// TIA Portal project "Can_Van_An_Modbus_ASCII" (V21)

(* hardware
DEVICE "S7-1500/ET200MP station_1"  S7-1500 station
   slot 0: "Rail_0"  Rack  6ES7 590-1***0-0AA0
   slot 1: "PLC_1"  CPU 1513-1 PN  6ES7 513-1AL02-0AB0  V2.9
      slot 3: "CPU display_1"  6ES7591-1AA00-0AA0
      slot 32768: "PROFINET interface_1"  X1
         slot 32769: "Port_1"  X1 P1
         slot 32770: "Port_2"  X1 P2
      slot 34817: "Virtual CP interface port_1"  Virtual CP interface port  Virtual CP interface port
DEVICE "ET 200SP station_1"  ET 200SP-Station
   slot 0: "Rack_0"  Rack  6ES5 710-8MAx1
   slot 0: "IO device_1"  IM 155-6 PN ST  6ES7 155-6AU01-0BN0  V4.2
   slot 1: "CM PtP_1"  CM PtP  6ES7 137-6AA01-0BA0  V2.0
      slot 1: "CM PtP_1"  CM PtP Sub
   slot 2: "Server module_1"  Server module  6ES7 193-6PA00-0AA0  V1.1
      slot 1: "Server module_1"  Server module
   slot 127: "BA 2xRJ45"  BA 2xRJ45  6ES7 193-6AR00-0AA0  V0.0
      slot 1: "Port_1"  X1 P1R  6ES7 193-6AR00-0AA0  V0.0
      slot 2: "Port_2"  X1 P2R  6ES7 193-6AR00-0AA0  V0.0
*)

// ===== PLC "PLC_1"  CPU 1513-1 PN =====

VAR_GLOBAL   // PLC tag table "1_Default tag table"
   "System_Byte" AT %MB1 : Byte;
   "FirstScan" AT %M1.0 : Bool;
   "DiagStatusUpdate" AT %M1.1 : Bool;
   "AlwaysTRUE" AT %M1.2 : Bool;
   "AlwaysFALSE" AT %M1.3 : Bool;
   "Clock_Byte" AT %MB0 : Byte;
   "Clock_10Hz" AT %M0.0 : Bool;
   "Clock_5Hz" AT %M0.1 : Bool;
   "Clock_2.5Hz" AT %M0.2 : Bool;
   "Clock_2Hz" AT %M0.3 : Bool;
   "Clock_1.25Hz" AT %M0.4 : Bool;
   "Clock_1Hz" AT %M0.5 : Bool;
   "Clock_0.625Hz" AT %M0.6 : Bool;
   "Clock_0.5Hz" AT %M0.7 : Bool;
END_VAR

VAR_GLOBAL   // PLC tag table "2_Bit_Tam(2-10)"
   "bTrigger1" AT %M2.0 : Bool;
   "bTrigger2" AT %M2.1 : Bool;
   "bTrigger3" AT %M2.2 : Bool;
   "bTrigger4" AT %M2.3 : Bool;
   "bTrigger5" AT %M2.4 : Bool;
   "bTrigger6" AT %M2.5 : Bool;
   "bTrigger7" AT %M2.6 : Bool;
   "bTrigger8" AT %M2.7 : Bool;
   "bTrigger9" AT %M3.0 : Bool;
   "bTrigger10" AT %M3.1 : Bool;
END_VAR

VAR_GLOBAL   // PLC tag table "3_DataNodeRed(100-200)"
   "diWeight" AT %MD100 : DInt;
   "wErrorCodeWeight" AT %MW104 : Word;
   "wStatusPLC" AT %MW106 : Word;
END_VAR

TYPE "typePortConfigSettings"
   STRUCT
      port : Int;
      protocol : Int;
      baud : Int;
      parity : Int;
      dataBis : Int;
      stopBits : Int;
      flowCntr : Int;
   END_STRUCT;
END_TYPE

TYPE "StartConditionReceive"
   STRUCT
      wStartCond : Word;
      wIdleTime : Word;
      StartChar : Byte;
   END_STRUCT;
END_TYPE

// folder: Common

TYPE "typeDiagnostics"
TITLE = typeDiagnostics
// Provides a structure for detailed diagnostics
   STRUCT
      status : Word;   // Status of the block or error identification when error occurred
      subfunctionStatus : DWord;   // Status or return value of called FBs, FCs and system blocks
      stateNumber : DInt;   // State in the state machine of the block where the error occurred
   END_STRUCT;
END_TYPE

// folder: LMQTT

TYPE "LMQTT_typeConnParam"
TITLE = LMQTT_typeConnParams
// Specifies connection parameters for the mqtt connection
   STRUCT
      hwId : Hw_Any;   // Hardware identifier of the interface. 0: interface is selected automatically
      connId : Conn_Ouc := 1;   // Unique connection identifier (1..4095)
      broker : String;   // Hostname or IP address of broker
      port : UInt := 1883;   // Port on the broker
      tls : Struct   // Parameters for TLS encryption
         enableTls : Bool;   // TRUE: Enables TLS, FALSE: disable TLS
         validateServerIdentity : Bool;   // TRUE: Validate server certificate, FALSE: No validation of server certificate
         brokerCert : UDInt;   // ID of the broker's certificate in TIA Portal
         clientCert : UDInt;   // ID of the client's certificate in TIA Portal
      END_STRUCT;
      keepAlive : UInt;   // Keepalive mechanism for MQTT in seconds. 0: disabled.
   END_STRUCT;
END_TYPE

// folder: typeDefinitions

TYPE "LModbusAscii_typeAsciiConfiguration"
TITLE = Parameter dataset to configure Modbus interface
// Parameter dataset to configure Modbus interface
   STRUCT
      baud : UInt := 6;   // Baud rate, default is 9600 (6), 19200 (7), see manual for other definitions
      parity : UInt := 2;   // Parity, default is even (2), odd (3) or none (1)
      modeInterfacePTP : USInt := 4;   // Serial interface mode, default is RS485 (4, Half duplex, two-wire mode), RS232 (0, FullDuplex)
      numberOfRetries : USInt := 3;   // Number of retries if a transmission error occurs, default is 3
      transmissionWatchdog : Time := T#5S;   // Response timeout duration, default is 5 s
   END_STRUCT;
END_TYPE

TYPE "LModbusAscii_typeDiagnostics"
TITLE = typeDiagnosticsTemplate
   STRUCT
      status : Word;   // Status of the block or error identification when error occurred
      stateNumber : DInt;   // State in the state machine of the block where the error occurred
      subFunctionStatus : Word;   // Status or return value of called FBs, FCs and system blocks
   END_STRUCT;
END_TYPE

// folder: (top level)

DATA_BLOCK "Data_StateSystem"   // DB1
{ S7_Optimized_Access := 'FALSE' }
VERSION : 0.1
   VAR
      "LED_PLC-S7-1500" : Struct
         "PLC-S7-1500" : Hw_Io := 50;
         Mode : Int := 1;
         Ret_Val : Word;
      END_STRUCT;
      ET200SP : Struct
         Device1 : Array[0..127] of Bool;
         RetVal : Int;
      END_STRUCT;
      bPLC_OFF : Bool;
      bPLC_Run : Bool;
      bPLC_Stop : Bool;
      bESP200_OK : Bool;
      bESP200_Fault : Bool;
      bESP200_LostConnect : Bool;
      bDonePortConfig : Bool;
      bErrorPortConfig : Bool;
      wStatusPortConfig : Word;
      "bDoneSend Config" : Bool;
      bErrorSendConfig : Bool;
      wStatusSendConfig : Word;
      bDoneReceiveConfig : Bool;
      bErrorReceiveConfig : Bool;
      wStatusReceiveConfig : Word;
      bDoneModbusKeli : Bool;
      bBusyModbusKeli : Bool;
      bErrorModbuskeli : Bool;
      ConditionReceive : Receive_Conditions;
   END_VAR
BEGIN
END_DATA_BLOCK

DATA_BLOCK "LMQTT_Client_EMQX_DB"   // DB2
{ S7_Optimized_Access := 'TRUE' }
AUTHOR : Siemens Industry Online Support
FAMILY : LMQTT
VERSION : 4.2
// stored: InstanceOfName LMQTT_Client
"LMQTT_Client"
BEGIN
END_DATA_BLOCK

DATA_BLOCK "KELI_ReadWeight_DB"   // DB3
{ S7_Optimized_Access := 'TRUE' }
VERSION : 1.0
// stored: InstanceOfName KELI_ReadWeight
"KELI_ReadWeight"
BEGIN
END_DATA_BLOCK

DATA_BLOCK "MQTT_Client"   // DB5
{ S7_Optimized_Access := 'FALSE' }
VERSION : 0.1
   VAR
      Inputs : Struct
         enable : Bool;
         publish : Bool;
         subscribe : Bool;
         unsubscribe : Bool;
         connParam : "LMQTT_typeConnParam";
         cleanSession : Bool;
         clientIdentifier : WString;
         username : WString;
         password : WString;
         willtopic : WString;
         willMsgLen : UInt;
         qos : USInt;
         retain : Bool;
         mqttTopic : WString;
         publishMsgLen : UDInt;
         timeOut : Time;
      END_STRUCT;
      Outputs : Struct
         valid : Bool;
         done : Bool;
         busy : Bool;
         error : Bool;
         status : Word;
         diagnostics : "typeDiagnostics";
         sessionPresent : Bool;
         receivedMsgStatus : USInt;
         receivedMsgDataLen : UDInt;
      END_STRUCT;
      InOut : Struct
         willMsgPayload : Array[0..7] of Byte;
         publishMsgPayload : Array[0..7] of Byte;
         receivedTopic : WString;
         receivedMsgPayload : Array[0..7] of Byte;
      END_STRUCT;
   END_VAR
BEGIN
   Inputs.connParam.hwId := 64;
END_DATA_BLOCK

DATA_BLOCK "Data_Server"   // DB11
{ S7_Optimized_Access := 'FALSE' }
VERSION : 0.1
   VAR
      MB_TCPIP : TCON_IP_v4;
   END_VAR
BEGIN
   MB_TCPIP.InterfaceId := 64;
   MB_TCPIP.ID := 1;
   MB_TCPIP.ConnectionType := 11;
   MB_TCPIP.ActiveEstablished := False;
   MB_TCPIP.RemoteAddress.ADDR[1] := 0;
   MB_TCPIP.RemoteAddress.ADDR[2] := 0;
   MB_TCPIP.RemoteAddress.ADDR[3] := 0;
   MB_TCPIP.RemoteAddress.ADDR[4] := 0;
   MB_TCPIP.RemotePort := 0;
   MB_TCPIP.LocalPort := 502;
END_DATA_BLOCK

DATA_BLOCK "Data_FrameKeli"   // DB13
{ S7_Optimized_Access := 'FALSE' }
VERSION : 0.1
   VAR
      ton : TON_TIME;
      WeightRAW_RX : String;
      ReadWeight_TX : Array[0..7] of Byte;
   END_VAR
BEGIN
   ReadWeight_TX[1] := 16#03;   // function
   ReadWeight_TX[0] := 16#02;   // address
   ReadWeight_TX[3] := 16#01;   // Thanh ghi băt đầu low
   ReadWeight_TX[2] := 16#00;   // Thanh ghi băt đầu high
   ReadWeight_TX[4] := 16#00;   // Thanh ghi kết thúc high
   ReadWeight_TX[5] := 16#04;   // Thanh ghi kết thúc low
   ReadWeight_TX[6] := 16#15;   // CRC16L
   ReadWeight_TX[7] := 16#FA;   // CRC16L
END_DATA_BLOCK

FUNCTION_BLOCK "KELI_ReadWeight"   // FB3, SCL
{ S7_Optimized_Access := 'TRUE' }
VERSION : 1.1
// ===============================================================================
//  KELI_ReadWeight - Đọc khối lượng GROSS của đầu cân KELI D2008 qua MODBUS (TF = 1)
//  PLC: S7-1200 / S7-1500 + module CM RS485 (Freeport, dùng Send_P2P / Receive_P2P)
// -------------------------------------------------------------------------------
//  CÀI ĐẶT ĐẦU CÂN: tF = 1 (MODBUS command), Adr = địa chỉ 1..247, bt = baudrate, jn = parity
//  CÀI ĐẶT CỔNG CM (Port configuration):
//    - Baudrate / parity / 8 data bit / 1 stop bit: giống đầu cân
//    - Message end (Receive): "Recognize end of message by line idle time"
//      (đầu cân nghỉ >= 4 ký tự sau mỗi khung -> CM báo đã nhận đủ khung)
// 
//  KHUNG TIN (theo manual D2008, mục MODBUS command mode):
//    Lệnh gửi (requestFrame, 8 byte):
//      [0] địa chỉ  [1] 16#03  [2] 16#00  [3] 16#01  [4] 16#00  [5] 16#04  [6] CRC low  [7] CRC high
//      ví dụ địa chỉ 1: 16#01 03 00 01 00 04 15 C9
//    Phản hồi bình thường (13 byte):
//      [0] địa chỉ  [1] 16#03  [2] 16#08 (= 8 byte dữ liệu)
//      [3] dấu: '0' (16#30) = dương, '-' = âm  [4..9] 6 chữ số ASCII (Data5..Data0)  [10] số chữ số thập phân
//      [11] CRC low  [12] CRC high
//      ví dụ 20.00 kg: '0' '0' '0' '2' '0' '0' '0' '2' -> weight = 2000, decimals = 2
//    Phản hồi lỗi (exception, 5 byte): [0] địa chỉ  [1] 16#83  [2] mã exception  [3] CRC L  [4] CRC H
// 
//  CRC16 MODBUS: giá trị đầu 16#FFFF, đa thức 16#A001, tính trên mọi byte trừ 2 byte CRC,
//    gửi byte thấp trước, byte cao sau.
// 
//  OUTPUT GIÁ TRỊ CÂN:
//    weight    : khối lượng dạng số nguyên, có dấu, KHÔNG có dấu thập phân (vd 2000)
//    decimals  : số chữ số sau dấu thập phân (vd 2  ->  khối lượng thật = 2000 / 10^2 = 20.00)
//    weightRaw : chuỗi 8 ký tự đầu cân gửi về, đúng nguyên bản (vd '00020002')
// 
//  status : 0 = BAD (lỗi), 1 = GOOD (đọc tốt), 2 = UNCERTAIN (chưa có giá trị / đang retry)
// 
//  TỰ KHỞI ĐỘNG LẠI: autoRestart = TRUE -> sau khi báo lỗi, FB chờ restartDelay rồi
//    tự chạy lại từ đầu, không cần sườn lên ở execute. restartCount đếm số lần tự chạy lại.
//    resetRestartCount (IN_OUT): SCADA/HMI ghi TRUE -> restartCount = 0, FB tự trả tag về FALSE.
//      Nối vào 1 tag Bool trong DB (vd "HMI".resetRestartCount_Can1), không nối hằng số.
// 
//  [V1.1] ĐO THỜI GIAN PHẢN HỒI CỦA ĐẦU CÂN (timer độ phân giải 1 ms):
//    Bắt đầu đếm : khi FB bắt đầu gửi lệnh xuống đầu cân (vào bước 20 - SEND)
//    Kết thúc    : khi CM báo đã nhận xong khung trả lời (Receive_P2P.NDR ở bước 30)
//    KHÔNG tính  : thời gian kiểm tra CRC và đổi ra số cân (bước 40)
//    responseTime   : kết quả dạng Time (vd T#45MS)
//    responseTimeMs : kết quả dạng số ms (vd 45) - tiện hiển thị trên HMI / SCADA
//    Chỉ cập nhật khi nhận được khung; timeout / lỗi gửi -> giữ giá trị lần đo gần nhất.
//    Mỗi lần retry đo lại từ đầu -> kết quả là thời gian của lần gửi nhận được trả lời.
//    Lưu ý: FB chỉ thấy NDR khi được gọi, nên kết quả có thể lớn hơn thực tế tối đa 1 chu kỳ quét.
// 
//  BẢNG MÃ LỖI (errorCode) - subStatus cho biết thêm chi tiết:
//    16#0000 ERR_NONE                không lỗi
//    16#8101 ERR_PARAM_ADDRESS       requestFrame[0] không thuộc 1..247   sub = địa chỉ nhập
//    16#8102 ERR_PARAM_FUNCTION      requestFrame[1] khác 16#03            sub = mã nhập
//    16#8103 ERR_PARAM_REGISTER      thanh ghi khác 16#0001 (gross)        sub = thanh ghi nhập
//    16#8104 ERR_PARAM_QUANTITY      số lượng khác 16#0004                 sub = số lượng nhập
//    16#8105 ERR_PARAM_CRC           sai CRC trong requestFrame            sub = CRC ĐÚNG (L H) để sửa
//    16#8201 ERR_RX_RESET            Receive_Reset lỗi                     sub = STATUS
//    16#8202 ERR_SEND                Send_P2P lỗi (truyền xuống)           sub = STATUS
//    16#8203 ERR_RECEIVE             Receive_P2P lỗi (nhận)                sub = STATUS
//    16#8204 ERR_TIMEOUT             không có phản hồi
//    16#8205 ERR_STATE_TIMEOUT       kẹt ở bước RX_RESET/SEND              sub = state
//    16#8301 ERR_FRAME_TOO_SHORT     gói ngắn hơn 5 byte                   sub = độ dài
//    16#8302 ERR_FRAME_ADDRESS       đầu cân khác trả lời                  sub = địa chỉ nhận
//    16#8303 ERR_FRAME_FUNCTION      mã hàm trả về sai                     sub = mã nhận
//    16#8304 ERR_FRAME_LENGTH        sai độ dài gói (phải 13 byte)         sub = độ dài
//    16#8305 ERR_FRAME_BYTE_COUNT    byte [2] khác 16#08                   sub = byte nhận
//    16#8401 ERR_CRC_MISMATCH        sai CRC gói nhận                      sub = CRC nhận (L H)
//    16#8501 ERR_EXCEPTION           đầu cân trả exception (16#83)         sub = mã exception
//    16#8601 ERR_WEIGHT_FORMAT       dấu / chữ số không hợp lệ             sub = vị trí byte lỗi
//    16#8602 ERR_WEIGHT_OVERLOAD     đầu cân báo quá tải (999999)
//    16#8603 ERR_DECIMAL_FORMAT      byte số thập phân không hợp lệ        sub = byte nhận
//    16#8701 ERR_UNDEFINED_STATE     lỗi state nội bộ                      sub = state
//    Có retry: 82xx, 83xx, 84xx. Không retry: 81xx, 85xx, 86xx, 8701.
// 
//  Bản 1 khối: CRC16 viết trực tiếp trong FB, không cần FC nào khác.
// 
//  LỊCH SỬ PHIÊN BẢN:
//    V1.0 (2026-10-07): bản đầu tiên - đọc gross weight, byte dấu '0' = dương,
//                       resetRestartCount dạng IN_OUT (FB tự trả về FALSE)
//    V1.1 (2026-10-08): thêm đo thời gian phản hồi của đầu cân
//                       (output responseTime, responseTimeMs; timer instResponseTimer)
// ===============================================================================
   VAR_INPUT
      execute : Bool;   // Sườn lên (0->1) = gửi 1 lệnh đọc
      hardwareId : Port;   // HW identifier của cổng RS485 trên CM
      requestFrame : Array[0..7] of Byte;   // Khung lệnh đọc gross: addr 03 00 01 00 04 CRC_L CRC_H
      timeout : Time := T#1S;   // Thời gian chờ phản hồi tối đa
      numberOfRetries : USInt := 2;   // Số lần gửi lại khi lỗi đường truyền/khung/CRC
      autoRestart : Bool := TRUE;   // TRUE = tự chạy lại sau khi báo lỗi
      restartDelay : Time := T#5S;   // Thời gian chờ trước khi tự chạy lại
   END_VAR
   VAR_OUTPUT
      done : Bool;   // TRUE = đọc thành công
      busy : Bool;   // TRUE = đang gửi / chờ phản hồi
      error : Bool;   // TRUE = lỗi (đã hết lượt retry)
      status : USInt := 2;   // 0 = BAD, 1 = GOOD, 2 = UNCERTAIN
      errorCode : Word;   // Mã lỗi, xem bảng ở đầu file
      subStatus : Word;   // Thông tin chi tiết của lỗi
      weight : DInt;   // Khối lượng số nguyên có dấu, không dấu thập phân
      decimals : USInt;   // Số chữ số thập phân (vị trí dấu '.' tính từ phải)
      weightRaw : String[8];   // 8 ký tự dữ liệu gốc: dấu + 6 số + số thập phân
      restartCount : UInt;   // Số lần FB đã tự chạy lại sau lỗi (chẩn đoán)
      responseTime : Time;   // [V1.1] Thời gian từ lúc gửi lệnh đến lúc nhận xong khung (vd T#45MS)
      responseTimeMs : DInt;   // [V1.1] Như responseTime nhưng dạng số ms (vd 45) cho HMI / SCADA
   END_VAR
   VAR_IN_OUT
      resetRestartCount : Bool;   // SCADA ghi TRUE = đưa restartCount về 0, FB tự trả về FALSE
   END_VAR
   VAR
      statState : Int;   // Bước hiện tại của state machine (0/10/20/30/40)
      statExecuteOld : Bool;   // Giá trị execute ở chu kỳ trước (bắt sườn lên)
      statDone : Bool;   // Bản trong của output done
      statBusy : Bool;   // Bản trong của output busy
      statError : Bool;   // Bản trong của output error
      statStatus : USInt := 2;   // Bản trong của output status
      statErrorCode : Word;   // Bản trong của output errorCode
      statSubStatus : Word;   // Bản trong của output subStatus
      statRetryCounter : USInt;   // Số lượt retry còn lại
      statTxBuffer : Array[0..7] of Byte;   // Khung gửi (chép từ requestFrame lúc bắt đầu lệnh)
      statTxLength : UInt := 8;   // Số byte cần gửi (= 8)
      statRxBuffer : Array[0..63] of Byte;   // Khung nhận từ đầu cân
      statRxLength : UInt;   // Số byte nhận được
      statCrcReceived : Word;   // CRC đầu cân gửi về, dạng (L H) (chẩn đoán)
      statCrcCalculated : Word;   // CRC PLC tự tính, dạng (L H) (chẩn đoán)
      statWeight : DInt;   // Bản trong của output weight
      statDecimals : USInt;   // Bản trong của output decimals
      statWeightRaw : String[8];   // Bản trong của output weightRaw
      instRxReset : Receive_Reset;   // Lệnh Siemens: xóa bộ đệm nhận của CM
      instSend : Send_P2P;   // Lệnh Siemens: gửi khung tin
      instReceive : Receive_P2P;   // Lệnh Siemens: nhận khung tin (kết thúc theo line idle)
      instTimeout : TON_TIME;   // Timer chờ phản hồi
      statRestartPending : Bool;   // TRUE = đã báo lỗi, đang chờ tự chạy lại
      statRestartCount : UInt;   // Bản trong của output restartCount
      instRestartTimer : TON_TIME;   // Timer đếm restartDelay trước khi tự chạy lại
      instStateWatchdog : TON_TIME;   // Timer canh bước RX_RESET / SEND không bị kẹt
      instResponseTimer : TON_TIME;   // [V1.1] Timer đo thời gian phản hồi (ET độ phân giải 1 ms)
      statResponseTime : Time;   // [V1.1] Bản trong của output responseTime
   END_VAR
   VAR_TEMP
      tempExecute : Bool;   // Bản sao execute trong chu kỳ này
      tempStartJob : Bool;   // TRUE = bắt đầu lệnh mới (sườn lên hoặc tự chạy lại)
      tempErrCode : Word;   // Mã lỗi phát hiện trong chu kỳ này
      tempSubStatus : Word;   // Chi tiết lỗi trong chu kỳ này
      tempRetryable : Bool;   // TRUE = lỗi này được phép gửi lại
      tempAddress : USInt;   // Địa chỉ đầu cân lấy từ requestFrame[0]
      tempRegister : Word;   // Thanh ghi bắt đầu trong requestFrame (byte 2..3)
      tempQuantity : Word;   // Số lượng thanh ghi trong requestFrame (byte 4..5)
      tempCrc : Word;   // CRC16 đang tính
      tempCrcLo : Byte;   // Byte thấp của CRC tính được
      tempCrcHi : Byte;   // Byte cao của CRC tính được
      tempBit : Int;   // Biến đếm 8 bit khi tính CRC
      tempLen : Int;   // Độ dài gói nhận
      tempIndex : Int;   // Biến đếm vòng FOR
      tempCode : USInt;   // Mã ASCII của ký tự đang xét
      tempValue : DInt;   // Giá trị cân đang ghép từ các chữ số
      tempNegative : Bool;   // TRUE = dấu '-'
      tempDigits : Int;   // Số chữ số đã đọc
      tempWeightOk : Bool;   // FALSE = gặp ký tự không hợp lệ
      tempBadIndex : Int;   // Vị trí byte lỗi (ghi vào subStatus)
      tempDecimals : USInt;   // Số chữ số thập phân đọc từ byte [10] các bước của state machine
   END_VAR
   VAR CONSTANT
      ST_IDLE : Int := 0;   // chờ lệnh
      ST_RX_RESET : Int := 10;   // xóa bộ đệm nhận
      ST_SEND : Int := 20;   // gửi lệnh
      ST_WAIT_RESPONSE : Int := 30;   // chờ phản hồi
      ST_PROCESS : Int := 40;   // phân tích gói nhận chất lượng dữ liệu (output status)
      QUALITY_BAD : USInt := 0;
      QUALITY_GOOD : USInt := 1;
      QUALITY_UNCERTAIN : USInt := 2;   // MODBUS
      FC_READ : Byte := 16#03;   // mã hàm đọc thanh ghi
      FC_EXCEPTION : Byte := 16#83;   // mã hàm báo lỗi (16#03 + 16#80)
      REG_GROSS : Word := 16#0001;   // thanh ghi gross weight
      QTY_GROSS : Word := 16#0004;   // đọc 4 thanh ghi = 8 byte dữ liệu
      BYTE_COUNT : Byte := 16#08;   // số byte dữ liệu trong phản hồi
      ADDRESS_MIN : USInt := 1;
      ADDRESS_MAX : USInt := 247;
      CRC_INIT : Word := 16#FFFF;   // giá trị đầu CRC16 MODBUS
      CRC_POLY : Word := 16#A001;   // đa thức CRC16 MODBUS (dạng đảo bit) độ dài khung (tính cả CRC)
      LEN_MIN_FRAME : Int := 5;   // khung exception
      LEN_WEIGHT_FRAME : Int := 13;   // khung giá trị cân
      RX_BUFFER_SIZE : Int := 64;
      RESPONSE_TIMER_PT : Time := T#1D;   // [V1.1] PT rất lớn: timer chỉ dùng ET để đo, không bao giờ chạy hết giờ
      OVERLOAD_VALUE : DInt := 999999;   // đầu cân báo quá tải
      DECIMALS_MAX : USInt := 5;   // 6 chữ số -> tối đa 5 số sau dấu '.' ký tự ASCII
      CHR_ZERO : Byte := 16#30;   // 0 (đầu cân gửi ở byte dấu khi giá trị dương)
      CHR_PLUS : Byte := 16#2B;   // +
      CHR_MINUS : Byte := 16#2D;   // -
      CHR_SPACE : Byte := 16#20;   // khoảng trắng mã lỗi (xem bảng ở đầu file)
      ERR_NONE : Word := 16#0000;
      ERR_PARAM_ADDRESS : Word := 16#8101;
      ERR_PARAM_FUNCTION : Word := 16#8102;
      ERR_PARAM_REGISTER : Word := 16#8103;
      ERR_PARAM_QUANTITY : Word := 16#8104;
      ERR_PARAM_CRC : Word := 16#8105;
      ERR_RX_RESET : Word := 16#8201;
      ERR_SEND : Word := 16#8202;
      ERR_RECEIVE : Word := 16#8203;
      ERR_TIMEOUT : Word := 16#8204;
      ERR_STATE_TIMEOUT : Word := 16#8205;
      ERR_FRAME_TOO_SHORT : Word := 16#8301;
      ERR_FRAME_ADDRESS : Word := 16#8302;
      ERR_FRAME_FUNCTION : Word := 16#8303;
      ERR_FRAME_LENGTH : Word := 16#8304;
      ERR_FRAME_BYTE_COUNT : Word := 16#8305;
      ERR_CRC_MISMATCH : Word := 16#8401;
      ERR_EXCEPTION : Word := 16#8501;
      ERR_WEIGHT_FORMAT : Word := 16#8601;
      ERR_WEIGHT_OVERLOAD : Word := 16#8602;
      ERR_DECIMAL_FORMAT : Word := 16#8603;
      ERR_UNDEFINED_STATE : Word := 16#8701;
   END_VAR
BEGIN

    REGION Khởi tạo biến tạm cho chu kỳ này
        // Biến Temp không giữ giá trị giữa các chu kỳ quét -> đặt lại mỗi lần FB chạy.
        // Mặc định: không lỗi. Đoạn nào phát hiện lỗi sẽ gán tempErrCode,
        // phần "Xử lý lỗi / retry" ở cuối FB sẽ xử lý chung.
        #tempExecute := #execute;
        #tempErrCode := #ERR_NONE;
        #tempSubStatus := 16#0000;
        #tempRetryable := FALSE;
    END_REGION

    REGION Tự khởi động lại sau lỗi / canh bước bị kẹt
        // Watchdog: bước xóa bộ đệm (RX_RESET) và bước gửi (SEND) bình thường xong rất nhanh.
        // Nếu kẹt lâu hơn 'timeout' (lệnh Siemens không báo DONE cũng không báo ERROR)
        // thì phần "Watchdog hết giờ" bên dưới sẽ báo lỗi 16#8205 để FB thoát ra.
        #instStateWatchdog(IN := #statState = #ST_RX_RESET OR #statState = #ST_SEND, PT := #timeout);

        // [V1.1] Timer đo thời gian phản hồi: IN = TRUE suốt bước 20 (SEND) và 30 (WAIT_RESPONSE).
        //   - Vào bước 20 (bắt đầu gửi lệnh)  -> IN 0 -> 1 -> timer bắt đầu đếm từ 0 ms
        //   - Bước 20 -> 30                    -> IN vẫn = 1 -> timer đếm tiếp, không bị reset
        //   - Rời bước 30 (sang 40 / retry 10 / về 0) -> IN = 0 -> ET về 0, sẵn sàng lần đo sau
        //   Giá trị ET được chốt lại ở bước 30 đúng lúc Receive_P2P báo NDR (xem REGION 30).
        #instResponseTimer(IN := #statState = #ST_SEND OR #statState = #ST_WAIT_RESPONSE, PT := #RESPONSE_TIMER_PT);

        // Tự chạy lại: khi đã báo lỗi (statRestartPending = TRUE) và FB đang ở IDLE,
        // timer đếm 'restartDelay'. Hết giờ -> coi như có lệnh mới, chạy lại từ đầu.
        #instRestartTimer(IN := #autoRestart AND #statRestartPending AND #statState = #ST_IDLE, PT := #restartDelay);

        // Bắt đầu lệnh mới khi: có sườn lên ở execute HOẶC timer tự chạy lại hết giờ
        #tempStartJob := (#tempExecute AND NOT #statExecuteOld) OR #instRestartTimer.Q;

        IF #tempStartJob AND #statState = #ST_IDLE THEN
            // đếm số lần tự chạy lại (để biết trên HMI đường truyền có hay lỗi không)
            IF #instRestartTimer.Q AND #statRestartCount < 65535 THEN
                #statRestartCount := #statRestartCount + 1;
            END_IF;
            #statRestartPending := FALSE;
            // đưa các lệnh truyền thông về trạng thái ban đầu (REQ = FALSE)
            // để lần gọi REQ = TRUE tiếp theo chắc chắn có sườn lên
            #instRxReset(REQ := FALSE, "PORT" := #hardwareId);
            #instSend(REQ := FALSE, "PORT" := #hardwareId, BUFFER := #statTxBuffer, LENGTH := #statTxLength);
            #instTimeout(IN := FALSE, PT := #timeout);
        END_IF;

        // Reset bộ đếm số lần tự chạy lại: SCADA ghi resetRestartCount = TRUE
        // -> restartCount = 0, rồi FB tự ghi resetRestartCount = FALSE (tag ở PLC tự nhả,
        // SCADA không cần ghi FALSE). Đặt sau đoạn tăng bộ đếm để lệnh reset luôn được ưu tiên.
        IF #resetRestartCount THEN
            #statRestartCount := 0;
            #resetRestartCount := FALSE;
        END_IF;
    END_REGION

    // ===== STATE MACHINE: mỗi chu kỳ chỉ chạy 1 nhánh theo giá trị statState =====
    CASE #statState OF
        #ST_IDLE:
            REGION 0 - IDLE: chờ lệnh, chép và kiểm tra khung gửi
                IF #tempStartJob THEN
                    // có lệnh mới -> xóa kết quả của lần trước
                    #statDone := FALSE;
                    #statError := FALSE;

                    // chép requestFrame vào buffer gửi của FB: nếu requestFrame bị đổi
                    // trong lúc đang chạy thì khung đang gửi / dùng để so sánh vẫn không đổi
                    FOR #tempIndex := 0 TO 7 DO
                        #statTxBuffer[#tempIndex] := #requestFrame[#tempIndex];
                    END_FOR;

                    // ghép 2 byte thành 1 Word: byte cao dịch trái 8 bit rồi OR byte thấp
                    // ví dụ 16#00, 16#01 -> 16#0001
                    #tempAddress := BYTE_TO_USINT(#statTxBuffer[0]);
                    #tempRegister := SHL(IN := BYTE_TO_WORD(#statTxBuffer[2]), N := 8) OR BYTE_TO_WORD(#statTxBuffer[3]);
                    #tempQuantity := SHL(IN := BYTE_TO_WORD(#statTxBuffer[4]), N := 8) OR BYTE_TO_WORD(#statTxBuffer[5]);

                    REGION Kiểm tra nội dung requestFrame
                        // Kiểm tra lần lượt, gặp lỗi đầu tiên thì dừng (chuỗi IF..ELSIF).
                        IF #tempAddress < #ADDRESS_MIN OR #tempAddress > #ADDRESS_MAX THEN
                            // địa chỉ MODBUS phải 1..247
                            #tempErrCode := #ERR_PARAM_ADDRESS;
                            #tempSubStatus := USINT_TO_WORD(#tempAddress);

                        ELSIF #statTxBuffer[1] <> #FC_READ THEN
                            // chỉ hỗ trợ mã hàm 16#03
                            #tempErrCode := #ERR_PARAM_FUNCTION;
                            #tempSubStatus := BYTE_TO_WORD(#statTxBuffer[1]);

                        ELSIF #tempRegister <> #REG_GROSS THEN
                            // FB này chỉ đọc gross weight (thanh ghi 16#0001)
                            #tempErrCode := #ERR_PARAM_REGISTER;
                            #tempSubStatus := #tempRegister;

                        ELSIF #tempQuantity <> #QTY_GROSS THEN
                            // gross weight cần đọc đúng 4 thanh ghi (8 byte)
                            #tempErrCode := #ERR_PARAM_QUANTITY;
                            #tempSubStatus := #tempQuantity;
                        END_IF;
                    END_REGION

                    REGION Kiểm tra CRC của requestFrame
                        IF #tempErrCode = #ERR_NONE THEN
                            // --- tính CRC16 MODBUS trên 6 byte đầu (byte 0..5) ---
                            #tempCrc := #CRC_INIT;
                            FOR #tempIndex := 0 TO 5 DO
                                // XOR byte dữ liệu vào 8 bit thấp của CRC
                                #tempCrc := #tempCrc XOR BYTE_TO_WORD(#statTxBuffer[#tempIndex]);
                                // xử lý 8 bit: bit thấp nhất = 1 -> dịch phải rồi XOR đa thức,
                                //              bit thấp nhất = 0 -> chỉ dịch phải
                                FOR #tempBit := 1 TO 8 DO
                                    IF (#tempCrc AND 16#0001) <> 16#0000 THEN
                                        #tempCrc := SHR(IN := #tempCrc, N := 1) XOR #CRC_POLY;
                                    ELSE
                                        #tempCrc := SHR(IN := #tempCrc, N := 1);
                                    END_IF;
                                END_FOR;
                            END_FOR;
                            #tempCrcLo := WORD_TO_BYTE(#tempCrc);                     // 8 bit thấp
                            #tempCrcHi := WORD_TO_BYTE(SHR(IN := #tempCrc, N := 8));  // 8 bit cao

                            // khung đúng: byte 6 = CRC low, byte 7 = CRC high
                            IF #statTxBuffer[6] <> #tempCrcLo OR #statTxBuffer[7] <> #tempCrcHi THEN
                                #tempErrCode := #ERR_PARAM_CRC;
                                // subStatus = CRC ĐÚNG theo thứ tự trong khung (L rồi H)
                                // ví dụ địa chỉ 1 -> 16#15C9 -> nhập byte 6 = 16#15, byte 7 = 16#C9
                                #tempSubStatus := SHL(IN := BYTE_TO_WORD(#tempCrcLo), N := 8) OR BYTE_TO_WORD(#tempCrcHi);
                            END_IF;
                        END_IF;
                    END_REGION

                    IF #tempErrCode = #ERR_NONE THEN
                        // khung hợp lệ -> nạp số lần retry, báo bận, chuyển sang bước xóa bộ đệm nhận
                        #statRetryCounter := #numberOfRetries;
                        #statBusy := TRUE;
                        #statState := #ST_RX_RESET;
                    END_IF;

                ELSIF NOT #tempExecute THEN
                    // done / error giữ TRUE chừng nào execute còn TRUE; execute = FALSE thì xóa
                    #statDone := FALSE;
                    #statError := FALSE;
                END_IF;
            END_REGION

        #ST_RX_RESET:
            REGION 10 - RX_RESET: xóa bộ đệm nhận của CM
                // Xóa rác / phản hồi cũ còn trong CM để gói nhận sau đó chắc chắn
                // là phản hồi của lệnh sắp gửi.
                #instRxReset(REQ := TRUE, "PORT" := #hardwareId);
                IF #instRxReset.DONE THEN
                    #instRxReset(REQ := FALSE, "PORT" := #hardwareId);     // hạ REQ cho lần sau
                    FILL_BLK(IN := 16#00, COUNT := 64, OUT => #statRxBuffer[0]); // xóa buffer nhận của FB
                    #statRxLength := 0;
                    #statState := #ST_SEND;
                ELSIF #instRxReset.ERROR THEN
                    #tempErrCode := #ERR_RX_RESET;                        // lỗi 16#8201
                    #tempSubStatus := #instRxReset.STATUS;                // mã lỗi Siemens
                    #tempRetryable := TRUE;
                    #instRxReset(REQ := FALSE, "PORT" := #hardwareId);
                END_IF;
            END_REGION

        #ST_SEND:
            REGION 20 - SEND: gửi khung lệnh xuống đầu cân
                // REQ giữ TRUE đến khi Send_P2P báo DONE hoặc ERROR
                #instSend(REQ := TRUE, "PORT" := #hardwareId, BUFFER := #statTxBuffer, LENGTH := #statTxLength);
                IF #instSend.DONE THEN
                    // gửi xong -> hạ REQ, reset timer timeout, chuyển sang chờ phản hồi
                    #instSend(REQ := FALSE, "PORT" := #hardwareId, BUFFER := #statTxBuffer, LENGTH := #statTxLength);
                    #instTimeout(IN := FALSE, PT := #timeout);
                    #statState := #ST_WAIT_RESPONSE;
                ELSIF #instSend.ERROR THEN
                    #tempErrCode := #ERR_SEND;                            // lỗi 16#8202
                    #tempSubStatus := #instSend.STATUS;
                    #tempRetryable := TRUE;
                    #instSend(REQ := FALSE, "PORT" := #hardwareId, BUFFER := #statTxBuffer, LENGTH := #statTxLength);
                END_IF;
            END_REGION

        #ST_WAIT_RESPONSE:
            REGION 30 - WAIT_RESPONSE: chờ phản hồi từ đầu cân
                // Receive_P2P báo NDR khi CM nhận xong 1 khung
                // (khung kết thúc khi đường truyền nghỉ - cấu hình 'line idle time' trong cổng CM).
                #instReceive("PORT" := #hardwareId, BUFFER := #statRxBuffer);
                #instTimeout(IN := TRUE, PT := #timeout);

                IF #instReceive.NDR THEN
                    // [V1.1] Chốt thời gian phản hồi NGAY khi nhận xong khung, trước khi phân tích:
                    //   gọi lại timer (IN vẫn TRUE) để ET được cập nhật đến đúng thời điểm này,
                    //   rồi lưu ET -> thời gian kiểm tra CRC / đổi ra số cân ở bước 40 không bị tính vào.
                    #instResponseTimer(IN := TRUE, PT := #RESPONSE_TIMER_PT);
                    #statResponseTime := #instResponseTimer.ET;

                    // đã nhận đủ 1 gói -> lưu độ dài, chuyển sang phân tích
                    #statRxLength := #instReceive.LENGTH;
                    #statState := #ST_PROCESS;
                ELSIF #instReceive.ERROR THEN
                    // CM báo lỗi nhận (parity, framing, tràn bộ đệm...)
                    #tempErrCode := #ERR_RECEIVE;                         // lỗi 16#8203
                    #tempSubStatus := #instReceive.STATUS;
                    #tempRetryable := TRUE;
                ELSIF #instTimeout.Q THEN
                    // hết thời gian mà chưa nhận được gói hoàn chỉnh
                    #tempErrCode := #ERR_TIMEOUT;                         // lỗi 16#8204
                    #tempRetryable := TRUE;
                END_IF;
            END_REGION

        #ST_PROCESS:
            REGION 40 - PROCESS: phân tích gói nhận
                #tempLen := UINT_TO_INT(#statRxLength);
                #tempRetryable := TRUE;   // mặc định: lỗi gói tin được gửi lại

                REGION Bước 1 - Kiểm tra độ dài tối thiểu
                    IF #tempLen < #LEN_MIN_FRAME THEN
                        // gói quá ngắn (ngắn hơn cả khung exception 5 byte)
                        #tempErrCode := #ERR_FRAME_TOO_SHORT;
                        #tempSubStatus := INT_TO_WORD(#tempLen);
                    ELSIF #tempLen > #RX_BUFFER_SIZE THEN
                        // gói dài hơn buffer
                        #tempErrCode := #ERR_FRAME_LENGTH;
                        #tempSubStatus := INT_TO_WORD(#tempLen);
                    END_IF;
                END_REGION

                REGION Bước 2 - Kiểm tra CRC gói nhận
                    // Kiểm tra CRC trước: CRC sai thì mọi byte khác trong gói đều không tin được
                    IF #tempErrCode = #ERR_NONE THEN
                        // --- tính CRC16 MODBUS trên byte 0 .. (len - 3), bỏ 2 byte CRC cuối ---
                        #tempCrc := #CRC_INIT;
                        FOR #tempIndex := 0 TO #tempLen - 3 DO
                            #tempCrc := #tempCrc XOR BYTE_TO_WORD(#statRxBuffer[#tempIndex]);
                            FOR #tempBit := 1 TO 8 DO
                                IF (#tempCrc AND 16#0001) <> 16#0000 THEN
                                    #tempCrc := SHR(IN := #tempCrc, N := 1) XOR #CRC_POLY;
                                ELSE
                                    #tempCrc := SHR(IN := #tempCrc, N := 1);
                                END_IF;
                            END_FOR;
                        END_FOR;
                        #tempCrcLo := WORD_TO_BYTE(#tempCrc);
                        #tempCrcHi := WORD_TO_BYTE(SHR(IN := #tempCrc, N := 8));

                        // lưu lại để xem khi chẩn đoán, dạng (L H) giống thứ tự trong khung
                        #statCrcCalculated := SHL(IN := BYTE_TO_WORD(#tempCrcLo), N := 8) OR BYTE_TO_WORD(#tempCrcHi);
                        #statCrcReceived := SHL(IN := BYTE_TO_WORD(#statRxBuffer[#tempLen - 2]), N := 8)
                                            OR BYTE_TO_WORD(#statRxBuffer[#tempLen - 1]);

                        IF #statCrcReceived <> #statCrcCalculated THEN
                            // gói bị nhiễu / hỏng trên đường truyền
                            #tempErrCode := #ERR_CRC_MISMATCH;
                            #tempSubStatus := #statCrcReceived;
                        END_IF;
                    END_IF;
                END_REGION

                REGION Bước 3 - Kiểm tra cấu trúc khung
                    // Kiểm tra lần lượt, gặp lỗi đầu tiên thì dừng (chuỗi IF..ELSIF).
                    IF #tempErrCode = #ERR_NONE THEN
                        IF #statRxBuffer[0] <> #statTxBuffer[0] THEN
                            // địa chỉ trả về phải trùng địa chỉ đã gửi
                            #tempErrCode := #ERR_FRAME_ADDRESS;
                            #tempSubStatus := BYTE_TO_WORD(#statRxBuffer[0]);

                        ELSIF #statRxBuffer[1] = #FC_EXCEPTION THEN
                            // đầu cân trả exception: không thực hiện được lệnh
                            // -> gửi lại cũng vô ích nên không retry
                            #tempErrCode := #ERR_EXCEPTION;
                            #tempSubStatus := BYTE_TO_WORD(#statRxBuffer[2]);   // mã exception
                            #tempRetryable := FALSE;

                        ELSIF #statRxBuffer[1] <> #FC_READ THEN
                            // mã hàm trả về phải là 16#03
                            #tempErrCode := #ERR_FRAME_FUNCTION;
                            #tempSubStatus := BYTE_TO_WORD(#statRxBuffer[1]);

                        ELSIF #tempLen <> #LEN_WEIGHT_FRAME THEN
                            // khung giá trị cân phải đúng 13 byte
                            #tempErrCode := #ERR_FRAME_LENGTH;
                            #tempSubStatus := INT_TO_WORD(#tempLen);

                        ELSIF #statRxBuffer[2] <> #BYTE_COUNT THEN
                            // byte [2] = số byte dữ liệu, phải là 8
                            #tempErrCode := #ERR_FRAME_BYTE_COUNT;
                            #tempSubStatus := BYTE_TO_WORD(#statRxBuffer[2]);
                        END_IF;
                    END_IF;
                END_REGION

                REGION Bước 4 - Tách giá trị cân
                    IF #tempErrCode = #ERR_NONE THEN
                        // từ đây trở đi là lỗi nội dung (gói đúng CRC) -> gửi lại cũng vô ích
                        #tempRetryable := FALSE;
                        #tempValue := 0;
                        #tempNegative := FALSE;
                        #tempDigits := 0;
                        #tempWeightOk := TRUE;
                        #tempBadIndex := 0;

                        // --- byte [3]: dấu ---
                        // Thực tế đầu cân gửi '0' (16#30) khi giá trị dương, '-' (16#2D) khi âm.
                        // Vẫn chấp nhận '+' (16#2B, theo manual) và ' ' (16#20) cho chắc.
                        IF #statRxBuffer[3] = #CHR_MINUS THEN
                            #tempNegative := TRUE;                          // '-' -> giá trị âm
                        ELSIF #statRxBuffer[3] <> #CHR_ZERO
                            AND #statRxBuffer[3] <> #CHR_PLUS
                            AND #statRxBuffer[3] <> #CHR_SPACE
                        THEN
                            #tempWeightOk := FALSE;                         // không phải '0', '+', '-', ' '
                            #tempBadIndex := 3;
                        END_IF;

                        // --- byte [4..9]: 6 chữ số ASCII, Data5 (hàng cao nhất) .. Data0 ---
                        // ví dụ "002000" -> 2000
                        IF #tempWeightOk THEN
                            FOR #tempIndex := 4 TO 9 DO
                                #tempCode := BYTE_TO_USINT(#statRxBuffer[#tempIndex]);
                                IF #tempCode >= 48 AND #tempCode <= 57 THEN
                                    // chữ số '0'..'9': ghép vào giá trị (dịch 1 hàng rồi cộng)
                                    #tempValue := #tempValue * 10 + USINT_TO_DINT(#tempCode - 48);
                                    #tempDigits := #tempDigits + 1;
                                ELSIF #tempCode = 32 AND #tempDigits = 0 THEN
                                    // khoảng trắng ở đầu -> bỏ qua
                                    ;
                                ELSE
                                    // ký tự không hợp lệ -> ghi vị trí, dừng đọc
                                    #tempWeightOk := FALSE;
                                    #tempBadIndex := #tempIndex;
                                    EXIT;
                                END_IF;
                            END_FOR;
                        END_IF;

                        // --- byte [10]: số chữ số thập phân ---
                        // manual cho ví dụ dạng ASCII ('2' = 16#32); chấp nhận cả dạng số (16#02)
                        #tempCode := BYTE_TO_USINT(#statRxBuffer[10]);
                        IF #tempCode >= 48 AND #tempCode <= 57 THEN
                            #tempDecimals := #tempCode - 48;                // '0'..'9' -> 0..9
                        ELSE
                            #tempDecimals := #tempCode;                     // đã là số
                        END_IF;

                        IF NOT #tempWeightOk OR #tempDigits = 0 THEN
                            // dấu sai, có ký tự lạ hoặc không có chữ số nào
                            #tempErrCode := #ERR_WEIGHT_FORMAT;
                            #tempSubStatus := INT_TO_WORD(#tempBadIndex);

                        ELSIF #tempDecimals > #DECIMALS_MAX THEN
                            // số thập phân phải 0..5
                            #tempErrCode := #ERR_DECIMAL_FORMAT;
                            #tempSubStatus := BYTE_TO_WORD(#statRxBuffer[10]);

                        ELSIF #tempValue = #OVERLOAD_VALUE THEN
                            // đầu cân gửi 999999 khi quá tải
                            #tempErrCode := #ERR_WEIGHT_OVERLOAD;

                        ELSE
                            // ===== ĐỌC THÀNH CÔNG =====
                            IF #tempNegative THEN
                                #tempValue := -#tempValue;
                            END_IF;
                            #statWeight := #tempValue;          // vd 2000 (không có dấu thập phân)
                            #statDecimals := #tempDecimals;     // vd 2    (-> 20.00)
                            // weightRaw: chép nguyên 8 byte dữ liệu [3..10] thành chuỗi, vd '00020002'
                            Chars_TO_Strg(Chars := #statRxBuffer,
                                          pChars := 3,
                                          Cnt := 8,
                                          Strg => #statWeightRaw);
                            #statDone := TRUE;
                            #statBusy := FALSE;
                            #statError := FALSE;
                            #statStatus := #QUALITY_GOOD;
                            #statErrorCode := #ERR_NONE;
                            #statSubStatus := 16#0000;
                            #statState := #ST_IDLE;   // quay về chờ lệnh tiếp theo
                        END_IF;
                    END_IF;
                END_REGION
            END_REGION

        ELSE
            // statState mang giá trị không có trong danh sách (không bình thường)
            #tempErrCode := #ERR_UNDEFINED_STATE;
            #tempSubStatus := INT_TO_WORD(#statState);
    END_CASE;

    REGION Watchdog hết giờ
        // FB kẹt ở RX_RESET hoặc SEND quá 'timeout' mà không có DONE/ERROR -> báo lỗi 16#8205,
        // hạ REQ của các lệnh để lần chạy lại có sườn lên mới.
        IF #tempErrCode = #ERR_NONE AND #instStateWatchdog.Q
            AND (#statState = #ST_RX_RESET OR #statState = #ST_SEND)
        THEN
            #tempErrCode := #ERR_STATE_TIMEOUT;
            #tempSubStatus := INT_TO_WORD(#statState);
            #tempRetryable := TRUE;
            #instRxReset(REQ := FALSE, "PORT" := #hardwareId);
            #instSend(REQ := FALSE, "PORT" := #hardwareId, BUFFER := #statTxBuffer, LENGTH := #statTxLength);
        END_IF;
    END_REGION

    REGION Xử lý lỗi / retry (dùng chung cho mọi bước)
        IF #tempErrCode <> #ERR_NONE THEN
            IF #tempRetryable AND #statRetryCounter > 0 THEN
                // còn lượt retry -> gửi lại từ bước xóa bộ đệm, chưa báo error ra ngoài
                #statRetryCounter := #statRetryCounter - 1;
                #instStateWatchdog(IN := FALSE, PT := #timeout);   // reset watchdog
                #statStatus := #QUALITY_UNCERTAIN;                  // giá trị chưa được xác nhận
                #statState := #ST_RX_RESET;
            ELSE
                // hết lượt retry hoặc lỗi không cho retry -> báo lỗi ra ngoài
                #statDone := FALSE;
                #statBusy := FALSE;
                #statError := TRUE;
                #statStatus := #QUALITY_BAD;
                #statErrorCode := #tempErrCode;
                #statSubStatus := #tempSubStatus;
                #statRestartPending := TRUE;                        // bật chờ tự chạy lại sau restartDelay
                #instStateWatchdog(IN := FALSE, PT := #timeout);   // reset watchdog
                #statState := #ST_IDLE;
            END_IF;
        END_IF;
    END_REGION

    // lưu execute của chu kỳ này để chu kỳ sau bắt sườn lên
    #statExecuteOld := #tempExecute;

    REGION Ghi output
        // ghi từ biến static ra output 1 lần ở cuối khối -> output luôn nhất quán
        #done := #statDone;
        #busy := #statBusy;
        #error := #statError;
        #status := #statStatus;
        #errorCode := #statErrorCode;
        #subStatus := #statSubStatus;
        #weight := #statWeight;         // khi lỗi vẫn giữ giá trị đúng gần nhất
        #decimals := #statDecimals;
        #weightRaw := #statWeightRaw;
        #restartCount := #statRestartCount;
        #responseTime := #statResponseTime;                    // [V1.1] thời gian phản hồi dạng Time
        #responseTimeMs := TIME_TO_DINT(#statResponseTime);   // [V1.1] đổi Time -> số ms (Time lưu nội bộ theo ms)
        ENO := NOT #statError;
    END_REGION
END_FUNCTION_BLOCK

ORGANIZATION_BLOCK "Main"   // OB1, LAD, ProgramCycle
TITLE = "Main Program Sweep (Cycle)"
{ S7_Optimized_Access := 'TRUE' }
VERSION : 0.1
   VAR_INPUT
      Initial_Call : Bool;   // Initial call of this OB
      Remanence : Bool;   // =True, if remanent data are available
   END_VAR
   VAR_TEMP   // added for the SCL form of the ladder/FBD networks
      _w1 : Bool;
   END_VAR
BEGIN

REGION Network 1: Check PLC S7 1500
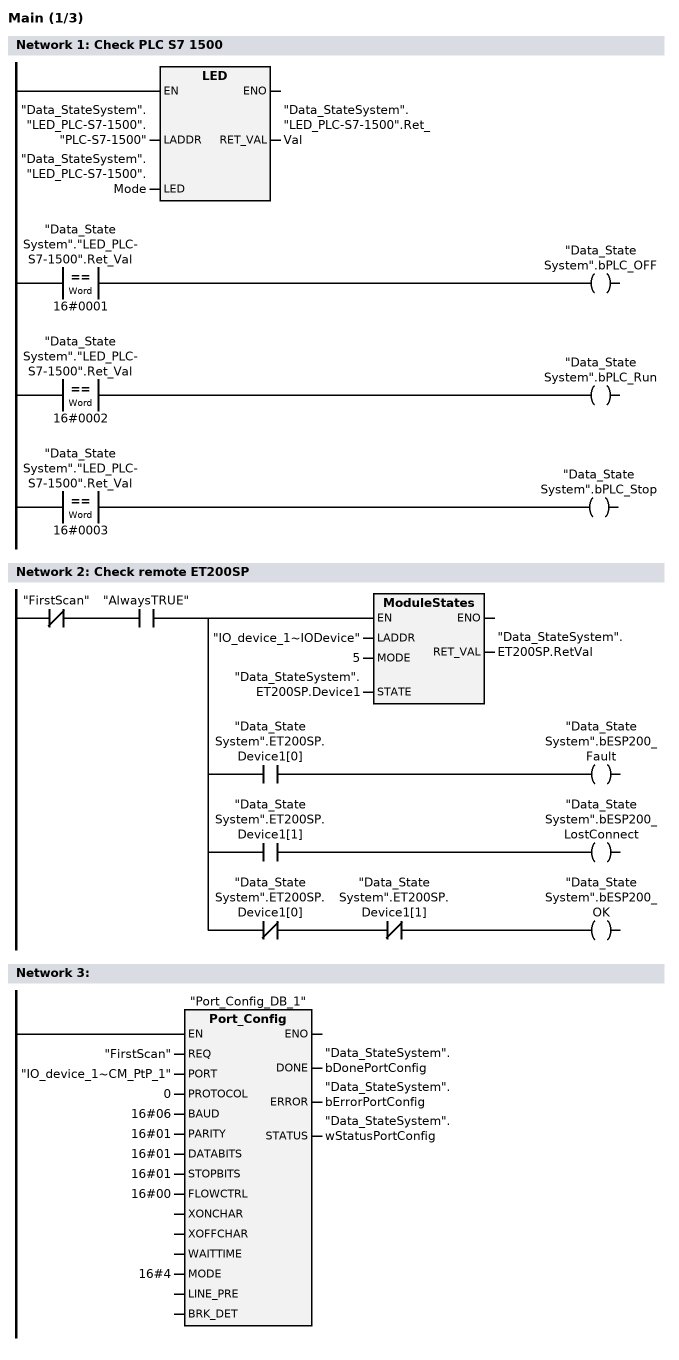
   "Data_StateSystem"."LED_PLC-S7-1500".Ret_Val := LED(LADDR := "Data_StateSystem"."LED_PLC-S7-1500"."PLC-S7-1500",
                           LED := "Data_StateSystem"."LED_PLC-S7-1500".Mode);
   "Data_StateSystem".bPLC_OFF := "Data_StateSystem"."LED_PLC-S7-1500".Ret_Val = 16#0001;
   "Data_StateSystem".bPLC_Run := "Data_StateSystem"."LED_PLC-S7-1500".Ret_Val = 16#0002;
   "Data_StateSystem".bPLC_Stop := "Data_StateSystem"."LED_PLC-S7-1500".Ret_Val = 16#0003;
END_REGION

REGION Network 2: Check remote ET200SP
   // no SCL statement known for ModuleStates: written as a call
   #_w1 := NOT "FirstScan" AND "AlwaysTRUE";
   IF #_w1 THEN
       "Data_StateSystem".ET200SP.RetVal := ModuleStates(LADDR := "IO_device_1~IODevice",
                               MODE := 5,
                               STATE := "Data_StateSystem".ET200SP.Device1);
   END_IF;
   "Data_StateSystem".bESP200_Fault := #_w1 AND "Data_StateSystem".ET200SP.Device1[0];
   "Data_StateSystem".bESP200_LostConnect := #_w1 AND "Data_StateSystem".ET200SP.Device1[1];
   "Data_StateSystem".bESP200_OK := #_w1 AND NOT "Data_StateSystem".ET200SP.Device1[0] AND NOT "Data_StateSystem".ET200SP.Device1[1];
END_REGION

REGION Network 3
   "Port_Config_DB_1"(REQ := "FirstScan",   // Port_Config
                      PORT := "IO_device_1~CM_PtP_1",
                      PROTOCOL := 0,
                      BAUD := 16#06,
                      PARITY := 16#01,
                      DATABITS := 16#01,
                      STOPBITS := 16#01,
                      FLOWCTRL := 16#00,
                      MODE := 16#4,
                      DONE => "Data_StateSystem".bDonePortConfig,
                      ERROR => "Data_StateSystem".bErrorPortConfig,
                      STATUS => "Data_StateSystem".wStatusPortConfig);
END_REGION

REGION Network 4
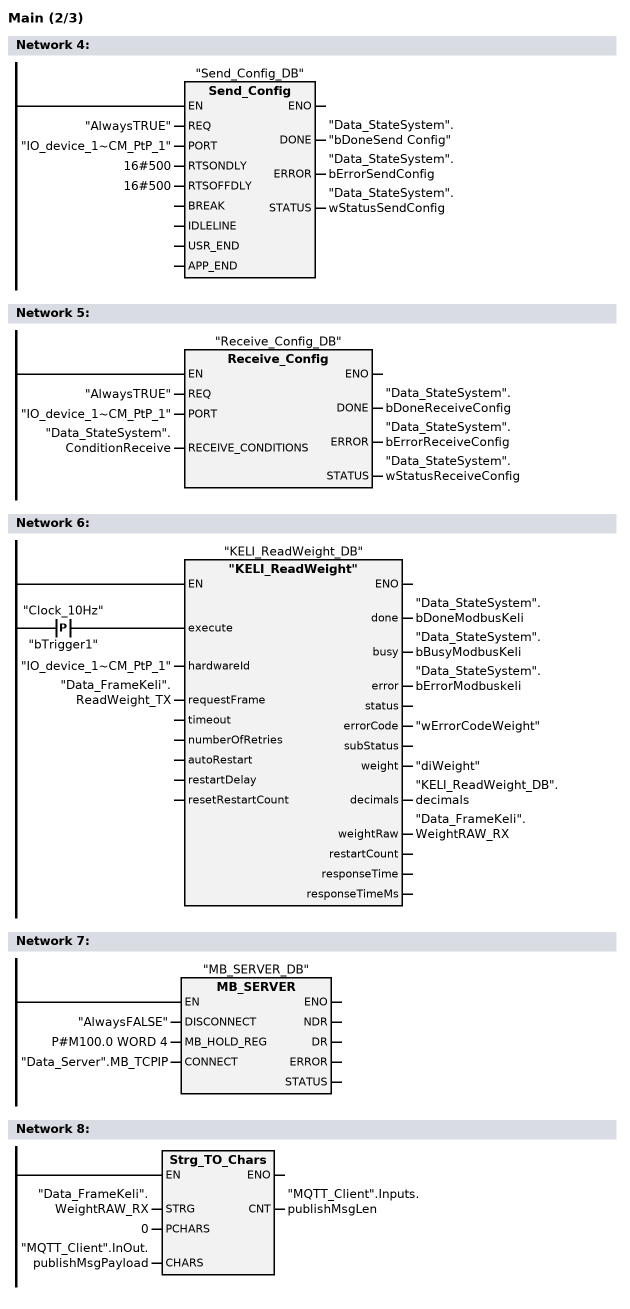
   "Send_Config_DB"(REQ := "AlwaysTRUE",   // Send_Config
                    PORT := "IO_device_1~CM_PtP_1",
                    RTSONDLY := 16#500,
                    RTSOFFDLY := 16#500,
                    DONE => "Data_StateSystem"."bDoneSend Config",
                    ERROR => "Data_StateSystem".bErrorSendConfig,
                    STATUS => "Data_StateSystem".wStatusSendConfig);
END_REGION

REGION Network 5
   "Receive_Config_DB"(REQ := "AlwaysTRUE",   // Receive_Config
                       PORT := "IO_device_1~CM_PtP_1",
                       Receive_Conditions := "Data_StateSystem".ConditionReceive,
                       DONE => "Data_StateSystem".bDoneReceiveConfig,
                       ERROR => "Data_StateSystem".bErrorReceiveConfig,
                       STATUS => "Data_StateSystem".wStatusReceiveConfig);
END_REGION

REGION Network 6
   RUNG wire#powerrail
      "KELI_ReadWeight_DB"(execute := wire#w1, hardwareId := "IO_device_1~CM_PtP_1", requestFrame := "Data_FrameKeli".ReadWeight_TX, timeout :=, numberOfRetries :=, autoRestart :=, restartDelay :=, resetRestartCount :=, done => "Data_StateSystem".bDoneModbusKeli, busy => "Data_StateSystem".bBusyModbusKeli, error => "Data_StateSystem".bErrorModbuskeli, status =>, errorCode => "wErrorCodeWeight", subStatus =>, weight => "diWeight", decimals => "KELI_ReadWeight_DB".decimals, weightRaw => "Data_FrameKeli".WeightRAW_RX, restartCount =>, responseTime =>, responseTimeMs =>)
   END_RUNG
   RUNG wire#powerrail
      P_Contact(operand := "Clock_10Hz", bit := "bTrigger1")
   END_RUNG wire#w1
   // the same network as SCL:
   #_w1 := "Clock_10Hz" AND NOT "bTrigger1";   // rising edge of "Clock_10Hz"
   "bTrigger1" := "Clock_10Hz";
   "KELI_ReadWeight_DB"(execute := #_w1,   // "KELI_ReadWeight"
                        hardwareId := "IO_device_1~CM_PtP_1",
                        requestFrame := "Data_FrameKeli".ReadWeight_TX,
                        done => "Data_StateSystem".bDoneModbusKeli,
                        busy => "Data_StateSystem".bBusyModbusKeli,
                        error => "Data_StateSystem".bErrorModbuskeli,
                        errorCode => "wErrorCodeWeight",
                        weight => "diWeight",
                        decimals => "KELI_ReadWeight_DB".decimals,
                        weightRaw => "Data_FrameKeli".WeightRAW_RX);
END_REGION

REGION Network 7
   "MB_SERVER_DB"(DISCONNECT := "AlwaysFALSE",   // MB_SERVER
                  MB_HOLD_REG := P#M100.0 WORD 4,
                  CONNECT := "Data_Server".MB_TCPIP);
END_REGION

REGION Network 8
   // no SCL statement known for Strg_TO_Chars: written as a call
   Strg_TO_Chars(Strg := "Data_FrameKeli".WeightRAW_RX,
                 pChars := 0,
                 Chars := "MQTT_Client".InOut.publishMsgPayload,
                 Cnt => "MQTT_Client".Inputs.publishMsgLen);
END_REGION

REGION Network 9
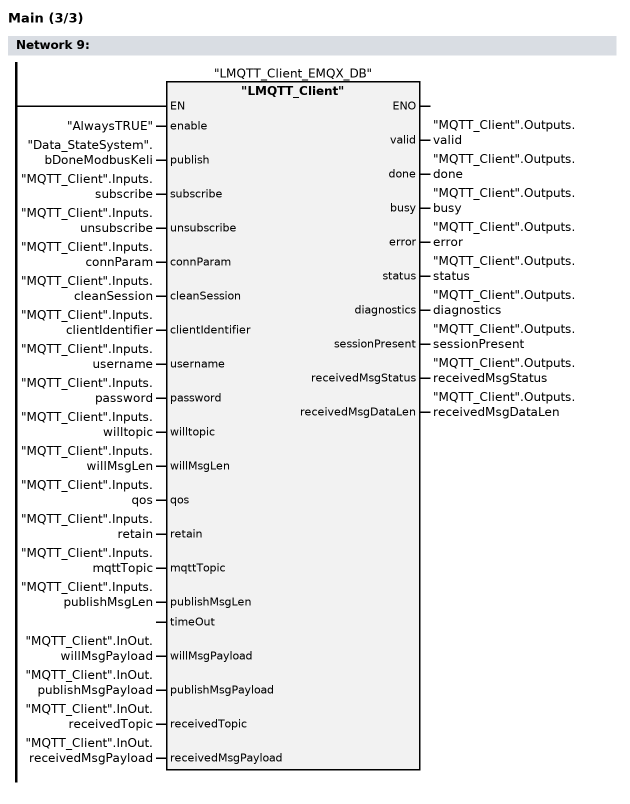
   RUNG wire#powerrail
      "LMQTT_Client_EMQX_DB"(enable := "AlwaysTRUE", publish := "Data_StateSystem".bDoneModbusKeli, subscribe := "MQTT_Client".Inputs.subscribe, unsubscribe := "MQTT_Client".Inputs.unsubscribe, connParam := "MQTT_Client".Inputs.connParam, cleanSession := "MQTT_Client".Inputs.cleanSession, clientIdentifier := "MQTT_Client".Inputs.clientIdentifier, username := "MQTT_Client".Inputs.username, password := "MQTT_Client".Inputs.password, willtopic := "MQTT_Client".Inputs.willtopic, willMsgLen := "MQTT_Client".Inputs.willMsgLen, qos := "MQTT_Client".Inputs.qos, retain := "MQTT_Client".Inputs.retain, mqttTopic := "MQTT_Client".Inputs.mqttTopic, publishMsgLen := "MQTT_Client".Inputs.publishMsgLen, timeOut :=, willMsgPayload := "MQTT_Client".InOut.willMsgPayload, publishMsgPayload := "MQTT_Client".InOut.publishMsgPayload, receivedTopic := "MQTT_Client".InOut.receivedTopic, receivedMsgPayload := "MQTT_Client".InOut.receivedMsgPayload, valid => "MQTT_Client".Outputs.valid, done => "MQTT_Client".Outputs.done, busy => "MQTT_Client".Outputs.busy, error => "MQTT_Client".Outputs.error, status => "MQTT_Client".Outputs.status, diagnostics => "MQTT_Client".Outputs.diagnostics, sessionPresent => "MQTT_Client".Outputs.sessionPresent, receivedMsgStatus => "MQTT_Client".Outputs.receivedMsgStatus, receivedMsgDataLen => "MQTT_Client".Outputs.receivedMsgDataLen)
   END_RUNG
   // the same network as SCL:
   "LMQTT_Client_EMQX_DB"(enable := "AlwaysTRUE",   // "LMQTT_Client"
                          publish := "Data_StateSystem".bDoneModbusKeli,
                          subscribe := "MQTT_Client".Inputs.subscribe,
                          unsubscribe := "MQTT_Client".Inputs.unsubscribe,
                          connParam := "MQTT_Client".Inputs.connParam,
                          cleanSession := "MQTT_Client".Inputs.cleanSession,
                          clientIdentifier := "MQTT_Client".Inputs.clientIdentifier,
                          username := "MQTT_Client".Inputs.username,
                          password := "MQTT_Client".Inputs.password,
                          willtopic := "MQTT_Client".Inputs.willtopic,
                          willMsgLen := "MQTT_Client".Inputs.willMsgLen,
                          qos := "MQTT_Client".Inputs.qos,
                          retain := "MQTT_Client".Inputs.retain,
                          mqttTopic := "MQTT_Client".Inputs.mqttTopic,
                          publishMsgLen := "MQTT_Client".Inputs.publishMsgLen,
                          willMsgPayload := "MQTT_Client".InOut.willMsgPayload,
                          publishMsgPayload := "MQTT_Client".InOut.publishMsgPayload,
                          receivedTopic := "MQTT_Client".InOut.receivedTopic,
                          receivedMsgPayload := "MQTT_Client".InOut.receivedMsgPayload,
                          valid => "MQTT_Client".Outputs.valid,
                          done => "MQTT_Client".Outputs.done,
                          busy => "MQTT_Client".Outputs.busy,
                          error => "MQTT_Client".Outputs.error,
                          status => "MQTT_Client".Outputs.status,
                          diagnostics => "MQTT_Client".Outputs.diagnostics,
                          sessionPresent => "MQTT_Client".Outputs.sessionPresent,
                          receivedMsgStatus => "MQTT_Client".Outputs.receivedMsgStatus,
                          receivedMsgDataLen => "MQTT_Client".Outputs.receivedMsgDataLen);
END_REGION
END_ORGANIZATION_BLOCK

// folder: Common

FUNCTION "IsIPAddress" : Bool   // FC1, SCL
TITLE = IsIPAddress
{ S7_Optimized_Access := 'TRUE' }
VERSION : 0.1
// Evaluates whether a given String contains a valid IP address
   VAR_INPUT
      address : String;   // Address to be evaluated
   END_VAR
   VAR_OUTPUT
      ipAddress : IP_V4;   // Parsed IP address if passed address is IP address
   END_VAR
   VAR_TEMP
      tempAddress : String;   // Passed address
      tempOctet : String;   // Current octet
      tempIndex : DInt;   // Index for loop
      tempPos : Int;   // Position of found separator
      tempNum : Int;   // Converted octet
      tempIp : IP_V4;   // Parsed IP address
   END_VAR
   // Ret_Val : Return value
   VAR CONSTANT
      MAX_VALUE : USInt := 255;   // Max. valid value of octet
      NUM_OCTETS : DInt := 4;   // Number of octets
      CHAR_ZERO : Char := '0';   // ASCII character '0'
   END_VAR
BEGIN
   REGION BLOCK INFO HEADER
     //===============================================================================
     // SIEMENS / (c)Copyright 2024
     //-------------------------------------------------------------------------------
     // Title:        IsIPAddress
     // Function:     Evaluates whether a given String contains a valid IP address
     // Library:      --
     // Author:       Siemens Industry Online Support
     // Tested with:  CPU 1515-2 PN V3.1
     // Engineering:  TIA Portal V17
     // Restrictions: --
     // Requirements: S7-1200 with firmware V4.4 or higher
     //               S7-1500 with firmware V2.0 or higher
     //-------------------------------------------------------------------------------
     // Change log table:
     // Version  | Date       | Expert in charge       | Changes applied
     //-------------------------------------------------------------------------------
     // 01.00.00 | 2024-02-12 | Online Support         | First released version
     //===============================================================================
   END_REGION

   #tempAddress := #address;
   #IsIPAddress := FALSE; // Will be overwritten if IP address is detected
   #ipAddress := #tempIp; // Zero output parameter

   FOR #tempIndex := 1 TO #NUM_OCTETS DO
     #tempPos := FIND(IN1 := #tempAddress, IN2 := '.'); // Find separator

     IF (#tempPos > 0 OR #tempIndex = #NUM_OCTETS) // Separator found with exception of last octet
       AND NOT (#tempPos > 0 AND #tempIndex = #NUM_OCTETS) // No separator found in last octet
       AND #tempPos <= 4 // 3  characters or less
     THEN
       IF #tempIndex < #NUM_OCTETS THEN // First three octets
         #tempOctet := LEFT(IN := #tempAddress, L := #tempPos - 1);
       ELSE// Last octet
         #tempOctet := #tempAddress;
       END_IF;

       STRG_VAL(IN := #tempOctet,
                FORMAT := 0,
                P := 1,
                OUT => #tempNum);

       IF #tempNum >= 0 AND #tempNum <= #MAX_VALUE // Within 0 and 255
         AND NOT (#tempNum = 0 AND #tempIndex = 1) // Not 0 in first octet
         AND NOT (#tempNum = 0 AND #tempOctet[1] <> #CHAR_ZERO) // Not 0 because of invalid character
       THEN
         #tempIp.ADDR[#tempIndex] := INT_TO_BYTE(#tempNum);
         #tempAddress := RIGHT(IN := #tempAddress, L := LEN(#tempAddress) - #tempPos); // Remove evaluated octet
       ELSE // Address is not IP address
         EXIT;
       END_IF;
     ELSE // Address is not IP address
       EXIT;
     END_IF;

     IF #tempIndex = #NUM_OCTETS THEN // End of loop reached, address is IP address
       #ipAddress := #tempIp;
       #IsIPAddress := true;
     END_IF;
   END_FOR;
END_FUNCTION

// folder: LMQTT

FUNCTION_BLOCK "LMQTT_Client"   // FB11, SCL
TITLE = LMQTT_Client
{ S7_Optimized_Access := 'TRUE' }
AUTHOR : Siemens Industry Online Support
FAMILY : LMQTT
VERSION : 4.2
// This block allows to connect to an MQTT Broker and publish data or receive data via a subscription.
   VAR_INPUT
      enable : Bool;   // Set TRUE, to establish a connection - set to FALSE to disconnect
      publish : Bool;   // Rising Edge: Sends a message
      subscribe : Bool;   // Rising Edge: Subscribes to a topic
      unsubscribe : Bool;   // Rising Edge: Unsubscribes to a topic
      connParam : "LMQTT_typeConnParam";   // Connection parameters
      cleanSession : Bool := TRUE;   // TRUE: Start a new session; FALSE: Session state must be saved by the broker
      clientIdentifier : WString;   // Client identifier
      username : WString;   // Username to connect
      password : WString;   // Password to connect
      willtopic : WString;   // Topic where the last will message is sent
      willMsgLen : UInt;   // Valid number of elements in Will Message Data Array. Max 65535 Byte allowed by MQTT Spec.
      qos : USInt;   // Quality of Service for publish/subscribe requests and last will. Subscribe only allows QoS 0 and 1
      retain : Bool;   // TRUE: Published Message will be set to retain on MQTT broker
      mqttTopic : WString;   // Mqtt Topic to Publish / Subscribe / Unsubscribe
      publishMsgLen : UDInt;   // Valid number of elements in publish message data Array
      timeOut : Time := T#5s;   // Sets the time out value for every request (publish/subscribe/unsubscribe/ping)
   END_VAR
   VAR_OUTPUT
      valid : Bool;   // TRUE: Valid set of output values available at the FB
      done : Bool;   // TRUE: If last Request was successfull
      busy : Bool;   // TRUE: FB is not finished and new output values can be expected
      error : Bool;   // TRUE: An error occurred during the execution of the FB
      status : Word := 16#7000;   // 16#0000 - 16#7FFF: Status of the FB, 16#8000 - 16#FFFF: Error identification
      diagnostics : "typeDiagnostics";   // Diagnostics information of FB
      sessionPresent : Bool;   // TRUE: A previous session was resumed; FALSE: New session established
      receivedMsgStatus : USInt;   // 0: No new Message, 1: New valid Message received and available at InOut area, 2: New message, but data is invalid (wrong message len or message could not be copied to InOut received topic or received message)
      receivedMsgDataLen : UDInt;   // Amount of Bytes received in receivedMessage INOUT area
   END_VAR
   VAR_IN_OUT
      willMsgPayload : Array[*] of Byte;   // Last will message Data - valid bytes in this array must be written in input 'willMsgLen'
      publishMsgPayload : Array[*] of Byte;   // Message Data to Publish - valid bytes in this array must be written in input 'publishMsgLen'
      receivedTopic : WString;   // Mqtt Topic of received message
      receivedMsgPayload : Array[*] of Byte;   // Mqtt message data that was received - valid bytes in this array indicated by 'receivedMsgDataLen' output
   END_VAR
   VAR
      statEnableOld : Bool;   // Old value of 'enable' input for edge detection
      statValid : Bool;   // Static value for output 'valid'
      statBusy : Bool;   // Static value for output 'busy'
      statError : Bool;   // Static value for output 'error'
      statErrorUserCleared : Bool;   // Error occurred that can only be solved by user; rising edge at enable input necessary
      statErrorAutoCleared : Bool;   // Error occurred that can be acknowledged by FB
      statStatus : Word := 16#7000;   // Static value for output 'status'
      statDone : Bool;   // Static value for output 'done'
      statRcvMsgStatus : USInt;   // Static value for output 'receivedMsgStatus'
      statRcvMsgDataLen : UDInt;   // Static value for output 'receivedMsgDataLen'
      statSubfunctionStatus : Word;   // Status or return value of called FBs, FCs and system blocks
      statFBErrorState : DInt;   // State in the state machine of the block where the error occurred
      statFBState : DInt := 0;   // State in the state machine of the FB
      statMqttConnectState : DInt := 0;   // State in the state machine of the MQTT Connection
      statMqttCommandState : DInt := 0;   // State in the state machine of the MQTT Commands when MQTT is connected
      statDisablingCompleted : Bool;   // TRUE: Disabling has been completed
      statEmptyDiagnostics : "typeDiagnostics";   // Empty diagnostics information (for initialization purposes only)
      statConnParam : Struct   // Connection parameters
         isQDN : Bool;   // QDN is used instead of IP address
         paramQDN : TCON_QDN_SEC;   // Parameter to assign QDN information
         paramIP : TCON_IP_V4_SEC;   // Parameter to assign IP information
      END_STRUCT;
      statSendBuffer : Array[0..#MAX_BUFFER_LEN_SEND] of Byte;   // Send buffer to send Data via TSend
      statRcvBuffer : Array[0..#MAX_BUFFER_LEN_RCV] of Byte;   // Receive buffer to receive Data via Trcv
      statRcvPayloadStorage : Array[0..#MAX_BUFFER_LEN_QOS2, 0..#MAX_BUFFER_LEN_RCV] of Byte;   // Buffer for storing the payload of received QoS 2 messages
      statRcvPacketIdStorage : Array[0..#MAX_BUFFER_LEN_QOS2] of Word;   // Buffer for storing the ID of received QoS 2 messages
      statRcvTopicStorage : Array[0..#MAX_BUFFER_LEN_QOS2] of WString;   // Buffer for storing the topic of received QoS 2 messages
      statRcvMsgPayloadLenStorage : Array[0..#MAX_BUFFER_LEN_QOS2] of UDInt;   // Buffer for storing the payload length of received QoS 2 messages
      statRcvTimestampStorage : Array[0..#MAX_BUFFER_LEN_QOS2] of DTL;   // Buffer for storing the time a QoS2 message arrived
      statPublishOld : Bool;   // Old value of 'publish' input for edge detection
      statSubscribeOld : Bool;   // Old value of 'subscribe' input for edge detection
      statUnsubscribeOld : Bool;   // Old value of 'unsubscribe' input for edge detection
      statTsendcReq : Bool;   // Static value to set send request
      statTsendcEnable : Bool;   // Static value to set tsend to enabled
      statTsendcLen : UDInt;   // Static value to len of tsend block
      statEnableTimerCommandWatchdog : Bool;   // Static value to start the command timer timeout
      statEnableMqttKeepAliveTimer : Bool;   // Static value to enable the Mqtt keepalive timer
      statMqttKeepAliveUsed : Bool;   // Static value to show if keepalive is used or deactivated
      statMqttKeepAliveTime : Time;   // Static value to store the keepalive Time interval
      statSendBufferPos : UInt;   // Static value to store the buffer position of the Tsend data area
      statPacketHeaderEncodeDone : Bool;   // Static value to show if a packet header was already encoded
      statSendPacketTotalRemLen : UDInt;   // Static value to store total packet length in bytes
      statEncodedRemPacketLenAsByte : Byte;   // Static value to store remaining length encoded as byte during calculation
      statUsernameLenUtf8Encoded : UInt;   // Static value to store total length of the username in utf8
      statPasswordLenUtf8Encoded : UInt;   // Static value to store total length of the password in utf8
      statWillTopicLenUtf8Encoded : UInt;   // Static value to store total length of the will topic in utf8
      statClientIdLenUtf8Encoded : UInt;   // Static value to store total length of the client id in utf8
      statWillQos : USInt;   // Static value to store the qos information of the will message
      statWillRetain : Bool;   // Static value to store the retain information of the will message
      statWillMessageCnt : UInt;   // Static value to store the amount of valid bytes in will message array
      statClientIdPos : DInt;   // Static value to store client id position during encoding
      statClientIdEncodeState : DInt;   // Static value to store the state during encoding
      statWillMessagePos : DInt;   // Static value to store will message position during encoding
      statWillMessageEncodeState : DInt;   // Static value to store the state during encoding
      statWillTopicPos : DInt;   // Static value to store will topic position during encoding
      statWillTopicEncodeState : DInt;   // Static value to store the state during encoding
      statUserNamePos : DInt;   // Static value to store user name position during encoding
      statUserNameEncodeState : DInt;   // Static value to store the state during encoding
      statPasswordPos : DInt;   // Static value to store password position during encoding
      statPasswordEncodeState : DInt;   // Static value to store the state during encoding
      statPacketId : UInt;   // Static value for the PacketId of each sent packet
      statPublishTopicLenUtf8Encoded : UInt;   // Static value to store total length of the publish topic in utf8
      statPublishQos : USInt;   // Static value to store the qos information of the publish message
      statPublishMessageCnt : UDInt;   // Static value to store the amount of valid bytes in publish message array
      statPublishTopicEncodeState : DInt;   // Static value to store the state during encoding
      statPublishTopicPos : DInt;   // Static value to store publish topic position during encoding
      statPacketIdEncoded : Bool;   // Static value to store if the packet id was encoded
      statPublishEncodeMessageState : DInt;   // Static value to store the state during encoding
      statPublishMessagePos : DInt;   // Static value to store publish message position during encoding
      statSubscribeQos : USInt;   // Static value to store the qos information of the subscribe message
      statSubscribeQosEncoded : Bool;   // Static value to store if the qos was encoded
      statSubscribeTopicPos : DInt;   // Static value to store subscribe topic position during encoding
      statSubscribeTopicEncodeState : DInt;   // Static value to store the state during encoding
      statSubscribeTopicLenUtf8Encoded : UInt;   // Static value to store total length of the subscribe topic in utf8
      statUnsubscribeTopicPos : DInt;   // Static value to store unsubscribe topic position during encoding
      statUnsubscribeTopicEncodeState : DInt;   // Static value to store the state during encoding
      statUnsubscribeTopicLenUtf8Encoded : UInt;   // Static value to store total length of the unsubscribe topic in utf8
      statRcvMsgQoS : UInt;   // Static value to store the qos information of the received message
      statRcvMsgTotalLen : UDInt;   // Static value to store the total len of the received message
      statRcvMsgTopicLen : UInt;   // Static value to store the total len of the received message topic
      statRcvMsgPayloadLen : UDInt;   // Static value to store the total len of the received message payload
      statRcvMsgPacketId : Word;   // Static value to store the packet id of the received message
      statRcvMsgTopicPos : DInt;   // Static value to store received message topic position during decoding
      statRcvMsgPayloadPos : DInt;   // Static value to store received message payload position during decoding
      statRcvMsgDecodeState : DInt;   // State in the state machine of the Rcv decoding
      statRcvMsgInternalStatus : USInt;   // Static value to store the internal status in case of topic or payload overflow
      statMqttPubRecRcv : USInt;   // Static value to store PUBREC of mqtt broker
      statMqttPubRelRcv : USInt;   // Static value to store PUBREL of mqtt broker
      statSendPubAckMsg : Bool;   // Static value to signal if PUBACK message must be sent
      statSendPubRecMsg : Bool;   // Static value to signal if PUBREC message must be sent
      statSendPubCompMsg : Bool;   // Static value to signal if PUBCOMP message must be sent
      statCommandInputOld : Bool;   // Static value used in ping exchange
      statCommandInputBackup : Byte;   // Static value used in ping exchange
      statRelPacketId : Word;   // Static value to store the ID of the message to be released
      statStoragePos : DInt;   // Static value to store the buffer index in which QoS 2 messages are stored
      statDecodedPayloadLenght : UDInt;   // Static value to store the last dataLen decoded
      statSessionPresent : Bool;   // Static value to store sessionPresent ouput
      instTsendC : TSEND_C;   // Tsend Instance
      instTrcv : TRCV;   // Trcv Instance
      instTimerCommandWatchdog : IEC_TIMER;   // Instance of the Timer for commands
      instMqttKeepAliveTimer : IEC_TIMER;   // Instance of the Timer for Mqtt keepalive
   END_VAR
   VAR_TEMP
      tempEnable : Bool;   // Temporary value for input 'enable'
      tempSubscribe : Bool;   // Temporary value for input 'subscribe'
      tempPublish : Bool;   // Temporary value for input 'publish'
      tempUnsubscribe : Bool;   // Temporary value for input 'unsubscribe'
      tempTsendcDone : Bool;   // Temporary value for instance of TsendC
      tempTsendcBusy : Bool;   // Temporary value for instance of TsendC
      tempTsendcError : Bool;   // Temporary value for instance of TsendC
      tempTsendcStatus : Word;   // Temporary value for instance of TsendC
      tempTrcvNdr : Bool;   // Temporary value for instance of Trcv
      tempTrcvBusy : Bool;   // Temporary value for instance of Trcv
      tempTrcvError : Bool;   // Temporary value for instance of Trcv
      tempTrcvStatus : Word;   // Temporary value for instance of Trcv
      tempTrcvRcvdLen : UDInt;   // Temporary value for instance of Trcv
      tempTrcvBufferPos : DInt;   // Temporary value for buffer position in trcv data array
      tempUserFlag : Bool;   // Temporary value to indicate if username is set
      tempPasswordFlag : Bool;   // Temporary value to indicate if passwordis set
      tempWillFlag : Bool;   // Temporary value to indicate if last will is set
      tempWillQoS1 : Bool;   // Temporary value to indicate if lastwill uses qos 1
      tempWillQoS2 : Bool;   // Temporary value to indicate if lastwill uses qos 2
      tempMaxWillMsgLen : DInt;   // Temporary value to store max will msg len
      tempLowerWillMsgArrayBoundary : DInt;   // Temporary value to store will msg data array lower bound from inout
      tempLoopCounter : DInt;   // Temporary value for several For loops
      tempBytesUsedUtf8 : USInt;   // Temporary value to store bytes used by a single character
      tempErrorConvertUtf8 : Bool;   // Temporary value to store if an error occured while converting character to utf8
      tempStatusConvertUtf8 : Word;   // Temporary value to store status code while converting character to utf8
      tempConvertedUtf8 : DWord;   // Temporary value to store the converted character in utf-8 format
      tempWordForSliceAddress : Word;   // Temporary value for several slice accesses
      tempCommandInput : Byte;   // Temporary value to set wether the command was publish subscribe or unsubscribe
      tempRcvMsgTypeCase : Byte;   // Temporary value to store which message type was received
      tempMaxPublishDataArrayLen : DInt;   // Temporary value to store the total length of the publish msg data array at inout
      tempMqttConnAckRcvStatus : USInt;   // Temporary value to store state of connection acknowledgement from broker
      tempMqttPingRspRcv : USInt;   // Temporary value to store PingResponse from broker
      tempMqttPubAckRcv : USInt;   // Temporary value to store Publish acknowledgement of mqtt broker
      tempMqttPubCompRcv : USInt;   // Temporary value to store Publish Completed of mqtt broker
      tempMqttSubAckRcv : USInt;   // Temporary value to store Subscribe acknowledgement of mqtt broker
      tempMqttUnSubAckRcv : USInt;   // Temporary value to store Unsubscribe acknowledgement of mqtt broker
      tempLowerBoundPublishDataArray : DInt;   // Temporary value to store lower bound of the publish data array
      tempMultiplierToDecode : UDInt;   // Temporary value to store the multiplier while packet decoding algorithm
      tempReceivedTopicStringMaxLen : DInt;   // Temporary value to store the max string len of the received topic
      tempReceivedMsgDataArrayTotalLen : DInt;   // Temporary value to store the total len of the received data msg array at inout
      tempUpperBoundRcvMsgDataArray : DInt;   // Temporary value to store the upper bound of the msg payload array
      tempReceivedTopic : WString;   // Temprary value to store received topic
      tempStorageIndex : UInt;   // Temporary value to store the index to access the QoS2 buffer
      tempCurrentTime : DTL;   // Temporary value to store current system time
      tempIntReturn : Int;   // Temporary value to store an Int return value
      tempTimeDiff : Time;   // Temporary value to calculate difference in time
   END_VAR
   VAR CONSTANT
      FB_STATE_NO_PROCESSING : DInt := 0;   // FB state: No processing
      FB_STATE_VALIDATE_INPUT : DInt := 10;   // FB state: Enabling - Validation of Inputs
      FB_STATE_TCP_CONNECTING : DInt := 20;   // FB state: Processing - TCP Connection establishing
      FB_STATE_OPERATING_MONITOR_TCP : DInt := 30;   // FB state: Processing - TCP Established, MQTT connection in progress
      FB_STATE_TCP_RECONNECTING : DInt := 40;   // FB state: Processing - TCP Connection must be re-established
      FB_STATE_DISABLING : DInt := 90;   // FB state: Disabling
      MQTT_CONNECT_STATE_NO_PROCESSING : DInt := 0;   // MQTT state: No processing
      MQTT_CONNECT_STATE_BUILD_PACKET : DInt := 100;   // MQTT state: Processing - build connect packet
      MQTT_CONNECT_STATE_SEND_PACKET_WAIT_FOR_CONNACK : DInt := 200;   // MQTT state: Processing - send connect packet
      MQTT_CONNECT_STATE_CONNECTED : DInt := 300;   // MQTT state: Processing - Connected to MQTT Broker
      MQTT_CONNECT_STATE_DISCONNECTED : DInt := 400;   // MQTT state: Processing - Disconnected to MQTT Broker
      MQTT_COMMAND_STATE_NO_PROCESSING : DInt := 0;   // MQTT Command state: No processing
      MQTT_COMMAND_STATE_BUILD_PUBLISH : DInt := 1;   // MQTT Command state: Build Publish packet
      MQTT_COMMAND_STATE_SEND_PUBLISH : DInt := 1000;   // MQTT Command state: Send Publish packet
      MQTT_COMMAND_STATE_BUILD_SUBSCRIBE : DInt := 2;   // MQTT Command state: Build Subscribe packet
      MQTT_COMMAND_STATE_SEND_SUBSCRIBE : DInt := 2000;   // MQTT Command state: Send Subscribe packet
      MQTT_COMMAND_STATE_BUILD_UNSUBSCRIBE : DInt := 4;   // MQTT Command state: Build Unsubscribe packet
      MQTT_COMMAND_STATE_SEND_UNSUBSCRIBE : DInt := 3000;   // MQTT Command state: Send Unsubscribe packet
      MQTT_COMMAND_STATE_SEND_PING : DInt := 8000;   // MQTT Command state: Send Ping packet
      MQTT_COMMAND_STATE_PING_RESP : DInt := 9000;   // MQTT Command state: Receive Ping packet
      STATUS_JOB_EXECUTED : Word := 16#0000;   // The last job was successfully executed
      STATUS_NO_CALL : Word := 16#7000;   // No job being currently processed
      STATUS_FIRST_CALL : Word := 16#7001;   // First call after incoming new job (rising edge 'enable')
      STATUS_SUBSEQUENT_CALL : Word := 16#7002;   // Subsequent call during active processing without further details
      STATUS_MQTT_CONNECTING : Word := 16#7003;   // Currently connecting to MQTT Broker
      STATUS_MQTT_CONNECTED : Word := 16#7004;   // Connected to MQTT Broker
      STATUS_MQTT_PING : Word := 16#7005;   // Processing Ping to Broker
      STATUS_MQTT_PUBLISH : Word := 16#7006;   // Processing Publish to Broker
      STATUS_MQTT_SUBSCRIBE : Word := 16#7008;   // Processing Subscribe to Broker
      STATUS_MQTT_UNSUBSCRIBE : Word := 16#7010;   // Processing Unsubscribe to Broker
      ERR_MQTT_COMMAND_MULTIPLE_INPUT : Word := 16#8001;   // Error - wrong operation - simultaneous input
      ERR_CLIENT_ID_NULL : Word := 16#8200;   // Error due to an incorrect client id at input
      ERR_CNT_EXCEEDS_ARRAY_DIMENSION : Word := 16#8210;   // Error due to an incorrect assignment of publish msg len or will msg len
      ERR_KEEPALIVE_INVALID : Word := 16#8220;   // Error due to an incorrect assignment of keepalive input
      ERR_QOS_INVALID : Word := 16#8230;   // Error due to an incorrect assignment of qos input
      ERR_MQTT_COMMAND_PUBLISH_TOPIC_INVALID : Word := 16#8300;   // Error - publish topic empty or invalid
      ERR_MQTT_COMMAND_SUBSCRIBE_TOPIC_INVALID : Word := 16#8310;   // Error - subscribe topic empty or invalid
      ERR_MQTT_COMMAND_UNSUBSCRIBE_TOPIC_INVALID : Word := 16#8320;   // Error - unsubscribe topic empty or invalid
      ERR_UNDEFINED_STATE : Word := 16#8600;   // Error due to an undefined state in state machine
      ERR_TCON_FAILED : Word := 16#8601;   // Error while trying to connect to mqtt broker with tcon
      ERR_TCON_TIMEOUT : Word := 16#8620;   // Error due to time out while trying to connect to broker
      ERR_MQTT_COMMAND_SEND_TIMEOUT : Word := 16#8650;   // Error - timeout while trying to sending data
      ERR_MQTT_CONNECT_TIMEOUT : Word := 16#8670;   // Error - timout while trying to connect via mqtt to broker
      ERR_MQTT_REM_LEN_INVALID : Word := 16#8700;   // Error due to receiving an invalid mqtt packet
      ERR_MQTT_MALFORMED_QOS_RECEIVED : Word := 16#8710;   // Error due to receiving an invalid mqtt packet
      ERR_MQTT_CONNACK_INVALID_SESSION_FLAG : Word := 16#8720;   // Error due to receiving an invalid mqtt packet
      ERR_MQTT_CONNACK_RETURN_CODE_INVALID : Word := 16#8730;   // Error due to receiving an invalid mqtt packet - see subfunction status for more information
      ERR_MQTT_PACKET_ID_INVALID : Word := 16#8740;   // Error due to receiving an invalid mqtt packet id
      ERR_MQTT_SUBACK_FAILURE : Word := 16#8750;   // Error because of failing to create a subscription
      ERR_CNT_QOS2_STORAGE_FULL : Word := 16#8760;   // Error due to the buffer of QoS 2 messages being full
      ERR_MSG_SKIPPED : Word := 16#8770;   // Error due to received message being skipped for not being fully inside the receive buffer
      ERR_TCP_RECONNECTING : Word := 16#9000;   // Error, lost connection to mqtt broker, reconnect ongoing
      MAX_BUFFER_LEN_RCV : UInt := 1459;   // Max. Buffer Len for TRCV
      MAX_BUFFER_LEN_SEND : UInt := 8191;   // Max. Buffer Len for TSEND on S7-1200/S7-1500
      MAX_BUFFER_LEN_QOS2 : UInt := 20;   // Max. Buffer Len for storing QoS 2 messages
      MAX_STORAGE_TIME_QOS2 : Time := T#10s;   // Max. Time that a QoS 2 message will be stored
      MAX_TOPIC_LEN_QOS2 : UInt := 254;   // Max. length of the topic string for QoS 2 messages
      EMPTY_BYTE : Byte := 16#00;   // Empty byte for initalisation
      EMPTY_WORD : Word;   // Empty word for initialization
      NO_COMMAND : Byte := 16#00;   // No Command for Executing Publish, Subscribe, Unsubscribe
      EMPTY_WSTRING : WString;   // Empty wstring for initalisation
      LEN_NULL : Int := 0;   // Integer 0 to compare length to zero
      INIT_UDINT_1 : UDInt := 1;   // Udint with value 1 for initalisation
      ARRAY_LEN_OFFSET_PLUS_1 : UInt := 1;   // Offset for array boundaries
      FIRST_CHARACTER : DInt := 1;   // First character in a character string
      ONE_DIMENSION : UDInt := 1;   // One dimensional array
      FIRST_ENCODING : DInt := 1;   // First encoding state while encoding messages
      SUBSEQUENT_ENCODING : DInt := 2;   // Followig encoding state while encoding messages if it takes multiple cycles
      ENCODE_DONE : DInt := 3;   // Last encoding state while encoding messages
      NOT_USED_NO_ENCODING : DInt := 5;   // No encoding state while encoding messages
      MSG_DECODE_STATE_NO_PROCESSING : DInt := 0;   // No message processing
      MSG_DECODE_STATE_TOPIC : DInt := 1;   // Message decoding state for topic
      MSG_DECODE_STATE_PACKET_ID_MSB : DInt := 2;   // Message decoding state for packet id msb
      MSG_DECODE_STATE_PACKET_ID_LSB : DInt := 3;   // Message decoding state for packet id lsb
      MSG_DECODE_STATE_PAYLOAD : DInt := 4;   // Message decoding state for packet payload
      MSG_DECODE_STATE_COMPLETED : DInt := 5;   // Message decoding state for packet decoded
      MSG_DECODE_STATUS_NO_NEW_MSG : USInt := 0;   // Message decoding status if no new message was received
      MSG_DECODE_STATUS_NEW_MSG_OK : USInt := 1;   // Message decoding status if a new message was received
      MSG_DECODE_STATUS_TOPIC_TOO_LONG : USInt := 2;   // Message decoding status if new message was received bute topic does not fit it inout topic (too shoirt)
      MSG_DECODE_STATUS_PAYLOAD_TOO_LONG : USInt := 2;   // Message decoding status if new message was received bute payload does not fit it inout payload(too shoirt)
      MQTT_QOS_0 : UInt := 0;   // Saving mqtt qos 0
      MQTT_QOS_1 : UInt := 1;   // Saving mqtt qos 1
      MQTT_QOS_2 : UInt := 2;   // Saving mqtt qos 2
      REMAINING_LEN_3 : Byte := 16#03;   // Remaining len in bytes is 3
      REMAINING_LEN_2 : Byte := 16#02;   // Remaining len in bytes is 2
      REMAINING_LEN_0 : Byte := 16#00;   // Remaining len in bytes is 0
      SUBSCRIBE_FAILURE : Byte := 16#80;   // Subscription failed flag.
      MQTT_NO_SESSION_PRESENT : Byte := 16#00;   // No session present indication
      KEEPALIVE_DISABLED : Time := T#0MS;   // Mqtt keepalive set to 0s
      TSENDC_JOB_DONE : Word := 16#0000;   // Status of tsendc if job was successful
      TSENDC_COM_CLOSED : Word := 16#0003;   // Status of tsendc if connection closed
      TSENDC_EST_OK : Word := 16#7004;   // Status of tsendc if connection ok
      TSENDC_DISCONNECTED : Word := 16#7000;   // Status of tsendc if disconnected from broker
      UINT_CONST_1000 : UInt := 1000;   // Calculation to seconds
      TWO_SECONDS : UInt := 2000;   // Calculation by 2 seconds
      THREE_SECONDS : UInt := 3;   // Upper limit is 3 seconds
      UTF_1_BYTE_USED : USInt := 1;   // If UTF uses 1 byte
      UTF_2_BYTE_USED : USInt := 2;   // If UTF uses 2 byte
      UTF_3_BYTE_USED : USInt := 3;   // If UTF uses 3 byte
      ONE_BYTE_LEN_INFO : UInt := 1;   // Adds one byte len info
      TWO_BYTE_LEN_INFO : UInt := 2;   // Adds two byte len info
      CONNECT_HEADER_10BYTE_LEN : UInt := 10;   // Connect header has always 10 byte minimum
      NO_RESPONSE : USInt := 0;   // If no response received from broker
      RESPONSE_GOOD : USInt := 1;   // If good response received from broker
      RESPONSE_PACKET_ID_INVALID : USInt := 2;   // If response received from broker but packet id invalid
      RESPONSE_SUBSCRIBE_FAILED : USInt := 3;   // If response received from broker but subscribption invalid
      MQTT_MSG_TYPE_CONNECT : Byte := 16#10;   // CONNECT MQTT Control Packet (see MQTT standard for more info)
      MQTT_MSG_TYPE_CONNACK : Byte := 16#20;   // CONNACK MQTT Control Packet (see MQTT standard for more info)
      MQTT_MSG_TYPE_PUBLISH : Byte := 16#30;   // PUBLISH MQTT Control Packet for QoS = 0 (see MQTT standard for more info)
      MQTT_MSG_TYPE_PUBACK : Byte := 16#40;   // PUBACK MQTT Control Packet (see MQTT standard for more info)
      MQTT_MSG_TYPE_PUBREC : Byte := 16#50;   // PUBREC MQTT Control Packet (see MQTT standard for more info)
      MQTT_MSG_TYPE_PUBREL : Byte := 16#60;   // PUBREL MQTT Control Packet (see MQTT standard for more info)
      MQTT_MSG_TYPE_PUBCOMP : Byte := 16#70;   // PUBCOM MQTT Control Packet (see MQTT standard for more info)
      MQTT_MSG_TYPE_SUBSCRIBE : Byte := 16#80;   // SUBSCRIBE MQTT Control Packet (see MQTT standard for more info)
      MQTT_MSG_TYPE_SUBACK : Byte := 16#90;   // SUBACK MQTT Control Packet (see MQTT standard for more info)
      MQTT_MSG_TYPE_UNSUBSCRIBE : Byte := 16#A0;   // UNSUBSCRIBE MQTT Control Packet (see MQTT standard for more info)
      MQTT_MSG_TYPE_UNSUBACK : Byte := 16#B0;   // UNSUBACK MQTT Control Packet (see MQTT standard for more info)
      MQTT_MSG_TYPE_PING : Byte := 16#C0;   // PING MQTT Control Packet (see MQTT standard for more info)
      MQTT_MSG_TYPE_PINGRESP : Byte := 16#D0;   // PINGRESP MQTT Control Packet (see MQTT standard for more info)
      MQTT_MSG_TYPE_DISCONNECT : Byte := 16#E0;   // DISCONNECT MQTT Control Packet (see MQTT standard for more info)
      MQTT_MSG_DECODING : Byte := 16#FF;   // STATE to show that currently a message is being decoded
      MQTT_MSG_QOS0 : Byte := 16#00;   // Bits for QoS 0 on the MQTT fixed header
      MQTT_MSG_QOS1 : Byte := 16#02;   // Bits for QoS 1 on the MQTT fixed header
      MQTT_MSG_QOS2 : Byte := 16#04;   // Bits for QoS 2 on the MQTT fixed header
      MQTT_MSG_QOS_BAD : Byte := 16#06;   // Bits for erroneous QoS on the MQTT fixed header
      BIT_MASK_HIGHBITS : Byte := 16#F0;   // MQTT Message Types only use High bits, so we only use High bits and ignore low bits
      BIT_MASK_QOS : Byte := 16#06;   // A Bit Mask to only validate recieved Byte against QOS Value
      MQTT_CONNACK_ACCEPTED : Byte := 16#00;   // Connect acknowledge flag in case no session present flag was not set
      DEFAULT_VALUE_ZERO : Int := 0;   // Default value for variables that are zero Based
      SEND_LEN_MULTIPLIER_UDINT_128 : UDInt := 128;   // Default mulitplier to calculate package length
      MAX_ALLOWED_PACKET_SIZE : UDInt := 2097152;   // The highest amount of payload to be sent by mqtt packet
      DEFAULT_MULTIPLIER_BYTE_127 : Byte := 16#7F;   // Default mulitplier to calculate package length
      CONN_PROTOCOL_NAME_0 : Byte := 16#00;   // Protocol version for mqtt
      CONN_PROTOCOL_NAME_4 : Byte := 16#04;   // Protocol version for mqtt
      CONN_PROTOCOL_MQTT_VERSION_3_1_1 : Byte := 16#04;   // Protocol version for mqtt
      BYTE_SIZE_CONNACK : USInt := 3;   // Size in bytes of a CONNACK packet (excluding header flags byte)
      BYTE_SIZE_PINGRESP : USInt := 1;   // Size in bytes of a PINGRESP packet (excluding header flags byte)
      BYTE_SIZE_PUBACK : USInt := 3;   // Size in bytes of a PUBACK packet (excluding header flags byte)
      BYTE_SIZE_PUBREC : USInt := 3;   // Size in bytes of a PUBREC packet (excluding header flags byte)
      BYTE_SIZE_PUBREL : USInt := 3;   // Size in bytes of a PUBREL packet (excluding header flags byte)
      BYTE_SIZE_PUBCOMP : USInt := 3;   // Size in bytes of a PUBCOMP packet (excluding header flags byte)
      BYTE_SIZE_SUBACK : USInt := 4;   // Size in bytes of a SUBACK packet (excluding header flags byte)
      BYTE_SIZE_UNSUBACK : USInt := 3;   // Size in bytes of a UNSUBACK packet (excluding header flags byte)
      BYTE_SIZE_PUBLISH : USInt := 6;   // Maximun size in bytes of the remaining length and topic length fields in a PUBLISH packet
   END_VAR
BEGIN
   REGION BLOCK INFO HEADER
       // ===============================================================================
       // SIEMENS (c)Copyright 2026
       // -------------------------------------------------------------------------------
       // Title:        LMQTT_Client
       // Function:     This FB implements an MQTT client. A user can publish data and
       //               subscribe to topics to receive data.
       // Library:      LMQTT
       // Author:       Siemens Industry Online Support
       // Tested with:  CPU 1516-3 PN/DP FW 2.9
       // Engineering:  TIA Portal V19
       // Restrictions: --
       // Requirements: S7-1200 with firmware V4.4 or higher
       //               S7-1500 with firmware V2.0 or higher
       // -------------------------------------------------------------------------------
       // Change log table:
       // Version  | Date       | Expert in charge   | Changes applied
       // ---------|------------|--------------------|------------------------------
       // 04.03.00 | 2026-08-12 | Online Support     | Added CleanSession flag
       //          |            |                    | Reordered interface
       // 04.02.00 | 2026-06-25 | Online Support     | Improved mechanism to deal with multiple messages arriving in the same PLC cycle
       // 04.01.02 | 2026-06-01 | Online Support     | Fixed bug when a timeout triggers at the same time a message arrives
       // 04.01.01 | 2026-02-11 | Online Support     | Fixed bug when receiving messages from subscriptions with QoS 2
       // 04.01.00 | 2024-10-28 | Online Support     | Fixed publishing OF more than 65535 messages (QoS > 0)
       //          |            |                    | Subscription with QoS2 implemented
       // 04.00.05 | 2024-06-05 | Online Support     | Fixed ActivateSecureConn reset
       // 04.00.04 | 2024-04-09 | Online Support     | Allowed lastWill without payload
       // 04.00.03 | 2024-02-12 | Online Support     | Improved evaluation of broker address
       // 04.00.02 | 2023-09-05 | Online Support     | Fixed bug that edge on publish/subscribe while PING is saved
       // 04.00.01 | 2023-08-30 | Online Support     | Fixed bug at TRCV and ConnID
       // 04.00.00 | 2023-08-04 | Online Support     | Broker can be addresses with hostname or IP address using one parameter
       //                                            | Reordered interface
       //                                            | Fixed bug at publish with QoS = 2
       // 03.00.05 | 2023-02-23 | Online Support     | Fixed bug that in rare situations no new commands were accepted
       // 03.00.04 | 2022-06-09 | Online Support     | Fixed bug that done was not set if input was reset
       // 03.00.03 | 2021-05-07 | Online Support     | Minor bug fixes
       // 03.00.00 | 2020-11-04 | Online Support     | New block interface with major improvements
       // 02.02.02 | 2020-03-16 | Online Support     | Improved issue with validateSubjectAlternateNameOfServer not setting correct bit
       // 02.02.01 | 2019-12-03 | Online Support     | Update to V16 and fusion with S7-1200 Lib
       // 02.01.00 | 2019-11-10 | Online Support     | Minor connection improvements. Updated some comments
       // 02.00.00 | 2018-06-04 | Online Support     | Added DNS support and Subscribe to topics
       // 01.00.00 | 2017-06-06 | Online Support     | First released version
       // ===============================================================================
   END_REGION

   #tempEnable := #enable; // Work with temporary value / create process image
   #tempPublish := #publish;  // Work with temporary value / create process image - only checked when MQTT is connected
   #tempSubscribe := #subscribe;  // Work with temporary value / create process image - only checked when MQTT is connected
   #tempUnsubscribe := #unsubscribe;  // Work with temporary value / create process image - only checked when MQTT is connected


   REGION OUC_BLOCK_CALLS
       // Only call if FB is processing
       IF #statStatus <> #STATUS_NO_CALL THEN
           // Connect and send
           IF #statConnParam.isQDN = TRUE THEN // Call if host is a domain name
               #instTsendC(REQ := #statTsendcReq,
                           CONT := #statTsendcEnable,
                           LEN := #statTsendcLen,
                           DONE => #tempTsendcDone,
                           BUSY => #tempTsendcBusy,
                           ERROR => #tempTsendcError,
                           STATUS => #tempTsendcStatus,
                           CONNECT := #statConnParam.paramQDN,
                           DATA := #statSendBuffer);
           ELSE
               #instTsendC(REQ := #statTsendcReq,
                           CONT := #statTsendcEnable,
                           LEN := #statTsendcLen,
                           DONE => #tempTsendcDone,
                           BUSY => #tempTsendcBusy,
                           ERROR => #tempTsendcError,
                           STATUS => #tempTsendcStatus,
                           CONNECT := #statConnParam.paramIP,
                           DATA := #statSendBuffer);
           END_IF;

           // Receive only when TCP operating
           #instTrcv(EN_R := (#statFBState = #FB_STATE_OPERATING_MONITOR_TCP),
                     ID := #statConnParam.paramQDN.ConnPara.ID,
                     ADHOC := true,
                     NDR => #tempTrcvNdr,
                     BUSY => #tempTrcvBusy,
                     ERROR => #tempTrcvError,
                     STATUS => #tempTrcvStatus,
                     RCVD_LEN => #tempTrcvRcvdLen,
                     DATA := #statRcvBuffer);

           // Monitor Time out
           #instTimerCommandWatchdog.TON(IN := #statEnableTimerCommandWatchdog,
                                         PT := #timeOut);
           // Mqtt Keepalive Timer
           #instMqttKeepAliveTimer.TON(IN := #statEnableMqttKeepAliveTimer,
                                       PT := #statMqttKeepAliveTime);
       END_IF;
   END_REGION

   REGION ENABLING/DISABLING_FUNCTION_BLOCK
       IF (#tempEnable = TRUE) AND (#statStatus = #STATUS_NO_CALL) THEN // Enable FB
           // First call; initialize FB
           #statValid := TRUE;
           #statBusy := TRUE;
           #statError := FALSE;
           #statDone := FALSE;
           #statErrorUserCleared := FALSE;
           #statErrorAutoCleared := FALSE;
           #statStatus := #STATUS_FIRST_CALL;
           #statSubfunctionStatus := #STATUS_JOB_EXECUTED;
           #statFBErrorState := 0;
           #diagnostics := #statEmptyDiagnostics;
           #statDisablingCompleted := FALSE;
           // State machine - start functionality
           #statFBState := #FB_STATE_VALIDATE_INPUT;

           // Initialize functionality: reset of variables, diagnostics, etc.
           #statPublishOld := FALSE;
           #statSubscribeOld := FALSE;
           #statUnsubscribeOld := FALSE;
           #statConnParam.isQDN := FALSE;
           #statTsendcReq := FALSE;
           #statTsendcEnable := FALSE;
           #statTsendcLen := 0;
           #statEnableTimerCommandWatchdog := FALSE;
           #statEnableMqttKeepAliveTimer := FALSE;
           #statMqttKeepAliveTime := #KEEPALIVE_DISABLED;
           #statMqttKeepAliveUsed := FALSE;
           #statSendBufferPos := 0;
           #statPacketHeaderEncodeDone := FALSE;
           #statSendPacketTotalRemLen := 0;
           #statEncodedRemPacketLenAsByte := #EMPTY_BYTE;
           #statClientIdPos := 0;
           #statClientIdEncodeState := 0;
           #statClientIdLenUtf8Encoded := 0;
           #statUserNamePos := 0;
           #statUserNameEncodeState := #FIRST_ENCODING;
           #statUsernameLenUtf8Encoded := 0;
           #statPasswordPos := 0;
           #statPasswordEncodeState := #FIRST_ENCODING;
           #statPasswordLenUtf8Encoded := 0;
           #statWillQos := 0;
           #statWillRetain := FALSE;
           #statWillMessageCnt := 0;
           #statWillMessagePos := 0;
           #statWillMessageEncodeState := #FIRST_ENCODING;
           #statWillTopicLenUtf8Encoded := 0;
           #statWillTopicPos := 0;
           #statWillTopicEncodeState := #FIRST_ENCODING;
           #statPacketId := 0;
           #statPublishTopicLenUtf8Encoded := 0;
           #statPublishQos := 0;
           #statPublishMessageCnt := 0;
           #statPublishTopicEncodeState := #FIRST_ENCODING;
           #statPublishTopicPos := 0;
           #statPacketIdEncoded := FALSE;
           #statPublishEncodeMessageState := #FIRST_ENCODING;
           #statPublishMessagePos := 0;
           #statSubscribeQos := 0;
           #statSubscribeQosEncoded := FALSE;
           #statSubscribeTopicPos := 0;
           #statSubscribeTopicEncodeState := #FIRST_ENCODING;
           #statSubscribeTopicLenUtf8Encoded := 0;
           #statUnsubscribeTopicPos := 0;
           #statUnsubscribeTopicEncodeState := #FIRST_ENCODING;
           #statUnsubscribeTopicLenUtf8Encoded := 0;
           #statRcvMsgQoS := 0;
           #statRcvMsgTotalLen := 0;
           #statRcvMsgTopicLen := 0;
           #statRcvMsgPayloadLen := 0;
           #statRcvMsgPacketId := 0;
           #statRcvMsgTopicPos := 0;
           #statRcvMsgPayloadPos := 0;
           #statRcvMsgDecodeState := #MSG_DECODE_STATE_NO_PROCESSING;
           #statRcvMsgInternalStatus := 0;
           #statRcvMsgStatus := 0;
           #statRcvMsgDataLen := 0;
           #statSendPubAckMsg := FALSE;
           #statSendPubRecMsg := FALSE;
           #statSendPubCompMsg := FALSE;
           #statStoragePos := 0;
           #statSessionPresent := FALSE;

           // Initialize functionality: call subsidiary FBs with FALSE
           FILL_BLK(IN := #EMPTY_BYTE,
                    COUNT := #MAX_BUFFER_LEN_SEND,
                    OUT => #statSendBuffer[0]);

           FILL_BLK(IN := #EMPTY_BYTE,
                    COUNT := #MAX_BUFFER_LEN_RCV,
                    OUT => #statRcvBuffer[0]);

           // Reset Packetid Buffer storage used by Subscribe QoS2 messages
           FILL_BLK(IN := #EMPTY_WORD,
                    COUNT := #MAX_BUFFER_LEN_QOS2,
                    OUT => #statRcvPacketIdStorage[0]);

           RESET_TIMER(#instTimerCommandWatchdog);
           RESET_TIMER(#instMqttKeepAliveTimer);

           // INIT SUB STATE MACHINES
           #statMqttConnectState := #MQTT_CONNECT_STATE_NO_PROCESSING;
           #statMqttCommandState := #MQTT_COMMAND_STATE_NO_PROCESSING;
           #statRcvMsgDecodeState := #MSG_DECODE_STATE_NO_PROCESSING;

